(* IEC 61131-3 sources: daoli-st-library/DL_Motion (part 8) *)

(* ---- FB_DL_AxisOverspeedGuard.st ---- *)
(*
  FB_DL_AxisOverspeedGuard  —  轴超速守卫（速度窗 + 加速度窗双判据） / Axis overspeed guard with velocity and acceleration windows
  分类 Category : DL_Motion
  版本 Version  : 1.0.0
  来源 Source   : t2-4-s7motion — 运动守卫族零检索深化
  溯源 Origin   : clean-room 实现，未复制任何源码行
  功能 Function : 1) 速度判据：|fVelocity| > fVelMax 持续 tVelTo → 故障级 03AC 独立锁存；
                  2) 加速度判据：离散差分 fAccEst := |v - vPrev| / tSamp（采样周期单位
                  已在头注释声明 [mm/s 每秒]），fAccEst > fAccMax 持续 tAccTo →
                  故障级 03AD 独立锁存（R190 归因唯一：两成因各自独立码位与独立出口）；
                  3) 故障解除式全当拍量（R240 落地），逐 BOOL 标注见段 5；
                  4) 速度回窗置信息级 04AB，加速度回窗置 04AC，使能沿置 04AD。
  边界 Boundary : ① 组态闸：fVelMax <= 0、fAccMax <= 0、tSamp <= 0、两超时 <= 0 → 03AB 锁存；
                  ② 差分分母下限 1.0E-6 s 防除零（TIME_TO_LREAL 后钳位）；
                  ③ 速度窗下限语义：判据为绝对值上窗，无下窗（下限 0 显式化）；
                  ④ 无 GVL 依赖：纯引脚输入输出，无外部变量引用，无物理 IO 地址。
  依赖 Depends  : I_DL_MotionAxis（注入，不实例化）；Standard.library（TON / R_TRIG）
  码表 Error codes（Motion 段 0004，窗口 03AB~03AD / 04AB~04AD）:
    16#0004_03AB 故障级：组态非法（速度窗/加速度窗/采样周期/超时域非法），锁存至 bReset
    16#0004_03AC 故障级：超速锁存（速度窗判据），锁存至 bReset
    16#0004_03AD 故障级：加速度超窗锁存（加速度窗判据），锁存至 bReset
    16#0004_04AB 信息级：速度恢复正常沿（回速度窗内）
    16#0004_04AC 信息级：加速度恢复正常沿（回加速度窗内）
    16#0004_04AD 信息级：守卫使能沿（bEnable 上升沿）
  修订历史 Revision :
    2026-11-19  v1.0.0  R41 首版（批次 2 · 序号 5）
*)

FUNCTION_BLOCK FB_DL_AxisOverspeedGuard
VAR_INPUT
    fVelMax      : REAL := 1000.0;    // 速度窗上限绝对值 [mm/s]，域 > 0 / Velocity window upper bound
    fAccMax      : REAL := 5000.0;    // 加速度窗上限 [mm/s²]，域 > 0 / Acceleration window bound
    tSamp        : TIME := T#10MS;    // 差分采样周期 [ms]，域 > 0 / Differentiation sample period
    tVelTo       : TIME := T#100MS;   // 超速确认超时 [ms]，域 > 0 / Overspeed confirm timeout
    tAccTo       : TIME := T#100MS;   // 超加速度确认超时 [ms]，域 > 0 / Over-acceleration confirm timeout
    bEnable      : BOOL := FALSE;     // 守卫使能 [-] / Guard enable
    bReset       : BOOL := FALSE;     // 复位，上升沿清故障锁存 / Reset edge clears fault latch
END_VAR
VAR_IN_OUT
    iAxis        : I_DL_MotionAxis;   // 运动轴引用（注入，不实例化）/ Motion axis reference
END_VAR
VAR_OUTPUT
    fVelAct      : REAL;              // 速度出口镜像 [mm/s] / Velocity outlet mirror
    fAccEst      : REAL;              // 加速度离散估计 [mm/s²] / Discrete acceleration estimate
    bVelFault    : BOOL;              // 超速独立锁存出口 [-] / Overspeed latch outlet
    bAccFault    : BOOL;              // 超加速度独立锁存出口 [-] / Over-acceleration latch outlet
    bFault       : BOOL;              // 聚合故障标志 [-] / Aggregate fault flag
    bError       : BOOL;              // 故障级标志（与聚合锁存同源）/ Fault flag
    nErrId       : UDINT;             // 事件码，0 = 无事件 / Event code
END_VAR
VAR
    tonVelTo     : TON;               // 超速确认定时器，无条件周期刷新 / Overspeed confirm timer
    tonAccTo     : TON;               // 超加速度确认定时器，无条件周期刷新 / Over-acceleration confirm timer
    rtReset      : R_TRIG;            // 复位沿实例，无条件刷新 / Reset edge instance
    rtEn         : R_TRIG;            // 使能沿实例，无条件刷新 / Enable edge instance
    _fVel        : REAL;              // 速度当拍量 [mm/s] / Current-scan velocity
    _fVelPrev    : REAL;              // 上拍速度快照 [mm/s] / Previous-scan velocity snapshot
    _fSampSec    : REAL;              // 生效采样周期 [s] / Effective sample period in seconds
    _bVelLat     : BOOL;              // 超速锁存位（锁存量）/ Overspeed latch bit
    _bAccLat     : BOOL;              // 超加速度锁存位（锁存量）/ Over-acceleration latch bit
    _bCfgBad     : BOOL;              // 组态非法锁存位（锁存量）/ Config-fault latch bit
    _uFault      : UDINT;             // 故障码锁存（锁存量）/ Latched fault code
    _uInfo       : UDINT;             // 信息码，每拍重算 / Transient info code
    _bVelOkPrev  : BOOL;              // 上拍速度窗内镜像（恢复沿判据）/ Previous velocity-in-window mirror
    _bAccOkPrev  : BOOL;              // 上拍加速度窗内镜像（恢复沿判据）/ Previous acceleration-in-window mirror
END_VAR

(* —— 段 0：定时器与沿实例无条件周期刷新（禁置于 IF/CASE 内） —— *)
_fVel := iAxis.fVelocity;                              // 速度当拍量
_fSampSec := TIME_TO_LREAL(tSamp) * 1.0E-3;            // 采样周期换算秒 [s]
IF _fSampSec < 1.0E-6 THEN
    _fSampSec := 1.0E-6;            // 差分分母下限防除零（下限钳位）
END_IF
fAccEst := ABS(_fVel - _fVelPrev) / _fSampSec;         // 加速度离散估计（差分口径）
rtReset(CLK := bReset);                                // 复位沿（每拍必调）
rtEn(CLK := bEnable);                                  // 使能沿（每拍必调）
tonVelTo(IN := bEnable AND (ABS(_fVel) > fVelMax), PT := tVelTo);   // 超速确认（每拍必调）
tonAccTo(IN := bEnable AND (fAccEst > fAccMax), PT := tAccTo);      // 超加速度确认（每拍必调）

(* —— 段 1：单拍量预清零（锁存量 _uFault/_bVelLat/_bAccLat/_bCfgBad 不入清单，禁同拍抹除） —— *)
_uInfo := 16#0000_0000;             // 信息码每拍重算
nErrId := 16#0000_0000;             // 事件码缺省无事件

(* —— 段 2：复位沿 + 组态域闸（当拍量判据） —— *)
IF rtReset.Q THEN                   // rtReset.Q = 当拍量
    _bVelLat := FALSE;              // 清超速锁存位
    _bAccLat := FALSE;              // 清超加速度锁存位
    _bCfgBad := FALSE;              // 清组态锁存位
    _uFault := 16#0000_0000;        // 清故障锁存码
END_IF
IF (fVelMax <= 0.0) OR (fAccMax <= 0.0) OR (TIME_TO_DINT(tSamp) <= 0)
   OR (TIME_TO_DINT(tVelTo) <= 0) OR (TIME_TO_DINT(tAccTo) <= 0) THEN
    _uFault := 16#0004_03AB;        // 故障级：组态非法
    _bCfgBad := TRUE;
END_IF

(* —— 段 3：双判据独立锁存（R190：速度/加速度归因唯一，各走独立码位与出口） —— *)
IF (NOT _bCfgBad) AND tonVelTo.Q THEN
    _uFault := 16#0004_03AC;        // 故障级：超速锁存
    _bVelLat := TRUE;
END_IF
IF (NOT _bCfgBad) AND tonAccTo.Q THEN
    _uFault := 16#0004_03AD;        // 故障级：加速度超窗锁存
    _bAccLat := TRUE;
END_IF

(* —— 段 4：故障解除式（R240 落地，逐 BOOL 标注）：
     rtReset.Q = 当拍量；ABS(_fVel) <= fVelMax = 当拍量；fAccEst <= fAccMax = 当拍量。
     均不含锁存量（_bVelLat/_bAccLat），解除边真实可达。 —— *)
IF rtReset.Q AND (NOT _bCfgBad) AND (ABS(_fVel) <= fVelMax) AND (fAccEst <= fAccMax) THEN
    _bVelLat := FALSE;              // 清超速锁存位（锁存量，仅此当拍量解除沿可清）
    _bAccLat := FALSE;              // 清超加速度锁存位（锁存量，同上）
    _uFault := 16#0000_0000;        // 清故障锁存码（锁存量，同上唯一解除路径）
END_IF

(* —— 段 5：信息码派生（当拍量判据） —— *)
IF (NOT _bCfgBad) AND bEnable THEN
    IF (ABS(_fVel) <= fVelMax) AND (NOT _bVelOkPrev) THEN
        _uInfo := 16#0004_04AB;     // 信息级：速度恢复沿
    END_IF
    IF (fAccEst <= fAccMax) AND (NOT _bAccOkPrev) THEN
        _uInfo := 16#0004_04AC;     // 信息级：加速度恢复沿（覆盖速度恢复沿，后到优先）
    END_IF
END_IF
IF rtEn.Q THEN
    _uInfo := 16#0004_04AD;         // 信息级：使能沿（使能优先报告）
END_IF

(* —— 段 6：出口单点映射（名实同源；锁存码回放，禁同拍抹除） —— *)
fVelAct := _fVel;                   // 速度出口镜像
bVelFault := _bVelLat OR _bCfgBad;  // 超速独立出口（组态非法并入聚合安全侧）
bAccFault := _bAccLat OR _bCfgBad;  // 超加速度独立出口（同上）
bFault := _bVelLat OR _bAccLat OR _bCfgBad;     // 聚合故障
IF bFault THEN
    nErrId := _uFault;              // 故障锁存码回放
ELSE
    nErrId := _uInfo;               // 信息码
END_IF
bError := bFault;                   // 故障标志与聚合锁存同源
_bVelOkPrev := (ABS(_fVel) <= fVelMax);   // 速度恢复沿判据快照
_bAccOkPrev := (fAccEst <= fAccMax);      // 加速度恢复沿判据快照
_fVelPrev := _fVel;                 // 上拍速度快照（段末统一写）

END_FUNCTION_BLOCK

(* ---- FB_DL_AxisPowerOnSelfTest.st ---- *)
(*==============================================================================
 * 组件名称 (Component)  : FB_DL_AxisPowerOnSelfTest
 * 所属子库 (Sublibrary) : DL_Motion
 * 当前版本 (Version)    : 1.0.1
 * 兼容性   (Platform)   : CODESYS 3.5 / TwinCAT 3 / 汇川 InoProShop / Machine Expert
 *                         仅依赖 Standard.library（TON / R_TRIG），零厂商方言
 * 来源标签 (Source)     : t2-4-s7motion（上电自检序列语义，clean-room 编写）
 * 功能描述 (Function)   : 轴上电自检五步序检：驱动就绪 -> 编码器回读（位置有效性
 *                         + 速率合理性）-> 限位状态巡检（常开 / 常闭组态域闸）->
 *                         驱动故障字扫描 -> 结论锁存。任一步失败即中止并禁使能
 *                         放行：bTestOk 出口供 FB_DL_SingleAxis 使能链消费。
 * 家族纪律 (R31)        : 不自造轴状态枚举——本件只消费快照与反馈引脚
 *                         （bDriveReady / fEncPos / fEncRate / 限位位 / 故障字），
 *                         轴状态机归运动层接口 I_DL_MotionAxis，本件零轴状态定义。
 * 边界与语义披露 (Boundary disclosure) :
 *   1) 步序超时逐段 TON 断输入（R40 家族口径）：步切换拍计时器复位一次
 *      （IN 串「步激活 AND NOT 步更替」），各步共用同一 tStepTimeout。
 *   2) 结论锁存：bTestOk 只在结论相置位并保持；解除 = 复位沿 AND 驱动就绪在位
 *      （终审两式：解除式可达，验收向量「复位沿 + 驱动就绪 -> 可重测」）。
 *   3) 限位组态域闸：nLimitMode 仅 0（常开）/ 1（常闭）合法，其余组态级故障；
 *      常闭口径下反馈 TRUE = 未压（健康），常开口径下反馈 TRUE = 被压。
 *   4) 上电即被压的限位按自检失败处置（轴未能验证自由行程，放行风险不可接受）。
 *   5) 编码器回读判据：位置 / 速率非有限（自反 + 差自减双判）或 |速率| 超
 *      fRateMax 均判步 2 失败（验收向量：回读 NaN -> 步 2 中止 bTestOk FALSE 置码）。
 *   6) 通用组态（速率上限 / 步超时）非法独立码位，与限位组态成因互异（R190）。
 * 故障码表 (Error codes) :
 *   16#0004_0363 [故障级] 步序超时（当前步 tStepTimeout 未达成）
 *                 反证：超时中止与「判据失败中止」eFault 输出组合相同，成因必须码位互异。
 *   16#0004_0364 [故障级] 编码器回读非法（位置 / 速率非有限或速率超合理域）
 *                 反证：步 2 中止与其它步中止输出组合相似，码位是唯一成因出口。
 *   16#0004_0365 [故障级] 限位组态模式非法（nLimitMode 非 0 / 1）
 *                 反证：限位步失败与编码器步失败输出组合相似，码位互异（R190）。
 *   16#0004_0366 [故障级] 上电限位被压（按生效接线口径判），自由行程未验证
 *                 反证：与组态非法同相中止但成因互异，码位独立。
 *   16#0004_0367 [故障级] 驱动故障字非零
 *                 反证：驱动故障字中止与编码器 / 限位 / 超时中止输出组合相似，成因互异码位独立。
 *   16#0004_0368 [故障级] 通用组态非法（速率上限 / 步超时域），拒绝启动
 *                 反证：拒绝启动与「未按触发」输出组合相同，码位唯一可见。
 * 码位总账 (Code ledger) : 16#0004_0363 / 0364 / 0365 / 0366 / 0367 / 0368 用
 * 依赖     (Depends)    : 无 DL_ 内部依赖；Standard.library: TON / R_TRIG
 * 红线自检 (Redline)    : R1 ✓ 零全局变量与 VAR_EXTERNAL ｜ R2 ✓ 零 %I/%Q 物理地址
 *                         R3 ✓ 纯 IEC 61131-3 ｜ R4 ✓ 非有限双判 / 域闸全枚举 / 码位 R45 配对
 *                         R5 ✓ 全变量中英双语同行注释 ｜ R6 ✓ 七态 ENUM + CASE + ELSE 兜底
 *                         R7 ✓ 三沿一计时主体最前部无条件刷新
 * 修订历史 (Revision)   :
 *   2026-11-22  v1.0.0  首版入库（R68 构建轮 · 批 3 · 目标 16）
 *   2026-11-22  v1.0.1  终审就地修①：组态锁存解除路径可达化（原 bCfgLatch 全文件零清零 -> 自检永久不可重测）
 *============================================================================*)

(*-----------------------------------------------------------------------------
 * 枚举: E_DL_SelfTestStep（归属 DL_Motion，与 FB_DL_AxisPowerOnSelfTest 同文件）
 * 说明: 本枚举是「自检步序」不是「轴状态」——轴状态归运动层接口（R31 家族纪律）。
 *----------------------------------------------------------------------------*)
TYPE E_DL_SelfTestStep :
(
    eIdle        := 0,    // 待触发：结论保持 / Idle, conclusion held
    eStDrive     := 10,   // 步 1：驱动就绪确认 / Step 1, drive ready
    eStEncoder   := 20,   // 步 2：编码器回读校验 / Step 2, encoder readback
    eStLimits    := 30,   // 步 3：限位状态巡检 / Step 3, limit switch patrol
    eStDriveWord := 40,   // 步 4：驱动故障字扫描 / Step 4, drive fault word scan
    eStConclude  := 50,   // 步 5：结论锁存 / Step 5, conclusion latch
    eFault       := 99    // 自检失败锁存：禁使能放行 / Self-test failed, enable release denied
);
END_TYPE

(*==============================================================================
 * 功能块: FB_DL_AxisPowerOnSelfTest
 * 调用约定: 每个扫描周期无条件调用一次；快照引脚须每拍刷新注入。
 *============================================================================*)
FUNCTION_BLOCK FB_DL_AxisPowerOnSelfTest
VAR_INPUT
    bTestTrig    : BOOL;                  // 自检触发（上升沿受理）/ Self-test trigger, rising edge
    bDriveReady  : BOOL;                  // 驱动就绪快照 / Drive ready snapshot
    fEncPos      : LREAL;                 // 编码器位置回读 [mm] / Encoder position readback [mm]
    fEncRate     : LREAL;                 // 编码器速率回读 [mm/s] / Encoder rate readback [mm per s]
    fRateMax     : LREAL := 100.0;        // 速率合理上限 [mm/s] / Plausible rate ceiling [mm per s]
    bLimitPosFb  : BOOL;                  // 正限位状态反馈（原始，TRUE = 电气有效）/ Positive limit feedback, raw
    bLimitNegFb  : BOOL;                  // 负限位状态反馈（原始）/ Negative limit feedback, raw
    nLimitMode   : INT   := 0;            // 限位接线模式：0 = 常开，1 = 常闭 / Wiring mode, 0 NO 1 NC
    uDriveFaultWord : WORD;               // 驱动故障字 / Drive fault word
    tStepTimeout : TIME  := T#2S;         // 单步超时 [s] / Step timeout [s]
    bEnable      : BOOL  := TRUE;         // 使能 / Enable
    bReset       : BOOL;                  // 上升沿：清结论与故障锁存（须驱动就绪在位）/ Rising edge: clear, drive ready required
END_VAR
VAR_OUTPUT
    bTestOk    : BOOL;                   // 自检结论：TRUE = 通过（锁存至复位 / 新测）/ Test passed, latched
    bTestDone  : BOOL;                   // 结论已出（通过或失败）/ Conclusion available
    bError     : BOOL;                   // 故障标志（自检失败 / 组态锁存归并）/ Fault flag merged
    uErrorId   : UDINT;                  // 故障码，0 = 无故障 / Error code, 0 = none
    eState     : E_DL_SelfTestStep;      // 当前步序（供 HMI 诊断）/ Current step for HMI diagnosis
END_VAR
VAR
    fbTrigTrig  : R_TRIG;                // 触发沿检测实例 / Trigger edge detector
    fbTrigReset : R_TRIG;                // 复位沿检测实例 / Reset edge detector
    tonStep     : TON;                   // 单步超时计时实例 / Step timeout timer
    eStateInt   : E_DL_SelfTestStep;     // 主状态机内部当前态 / Internal state machine state
    eStepPrev   : E_DL_SelfTestStep;     // 上拍步序快照（步更替判据）/ Previous step snapshot
    bStepActive : BOOL;                  // 当前步处于计时激活域 / Current step in the timed set
    bStepNew    : BOOL;                  // 本拍发生步更替（计时复位点）/ Step changed this scan
    bLimPosTrip : BOOL;                  // 按接线口径判的正限位被压 / Positive limit tripped per wiring
    bLimNegTrip : BOOL;                  // 负限位被压 / Negative limit tripped
    bEncBad     : BOOL;                  // 编码器回读非法 / Encoder readback illegal
    bCfgBad     : BOOL;                  // 本拍通用组态非法 / General config illegal
    bCfgLatch   : BOOL;                  // 通用组态锁存 / General config latch
    bModeBad    : BOOL;                  // 限位接线模式非法 / Wiring mode illegal
    bPassedInt  : BOOL;                  // 通过结论锁存内部副本 / Internal passed latch
    bDoneInt    : BOOL;                  // 结论已出锁存内部副本 / Internal done latch
    bErrorInt   : BOOL;                  // 本拍故障置位累加（出口归并）/ Fault set accumulator
    bFirstScan  : BOOL := TRUE;          // 上电首扫标志 / First-scan flag
END_VAR
VAR CONSTANT
    DL_ST_FIN_LIM   : LREAL := 1.0E30;   // LREAL 有限幅值判界 / LREAL finiteness bound
    DL_ST_MODE_NO   : INT   := 0;        // 常开接线模式号 / Normally-open mode id
    DL_ST_MODE_NC   : INT   := 1;        // 常闭接线模式号 / Normally-closed mode id
END_VAR

(*------------------------------------------------------------------------------
 * 段 1｜无条件刷新区（红线 R7）：二沿一计时主体最前部
 *      Unconditional refresh: two edges and one timer at the very top
 *      步更替拍计时复位一次（IN 串「步激活 AND NOT 步更替」，逐段断输入 R40）
 *-----------------------------------------------------------------------------*)
fbTrigTrig(CLK := bTestTrig);
fbTrigReset(CLK := bReset);

bStepNew := (eStateInt <> eStepPrev);

bStepActive := (eStateInt = E_DL_SelfTestStep.eStDrive)
               OR (eStateInt = E_DL_SelfTestStep.eStEncoder)
               OR (eStateInt = E_DL_SelfTestStep.eStLimits)
               OR (eStateInt = E_DL_SelfTestStep.eStDriveWord);

tonStep(IN := bStepActive AND (NOT bStepNew), PT := tStepTimeout);

(*------------------------------------------------------------------------------
 * 段 2｜上电首扫：结论与状态落安全侧（未测 = 不放行）
 *      First-scan init: conclusion to the safe side, untested means no release
 *-----------------------------------------------------------------------------*)
IF bFirstScan THEN
    eStateInt  := E_DL_SelfTestStep.eIdle;
    eStepPrev  := eStateInt;
    bPassedInt := FALSE;
    bDoneInt   := FALSE;
    bFirstScan := FALSE;
END_IF

(*------------------------------------------------------------------------------
 * 段 3｜每拍预清（FB32-1）：单拍标志，禁入锁存 / 快照
 *      Per-scan preset: single-scan flags only
 *-----------------------------------------------------------------------------*)
bErrorInt := FALSE;

(*------------------------------------------------------------------------------
 * 段 4｜组态域闸（R151 全枚举）：通用组态 + 限位接线模式（独立成因独立码 R190）
 *      Config gates: general config plus the wiring mode, distinct codes
 *      解除路径（R152 自证）：复位沿 AND 驱动就绪 AND 组态改对
 *-----------------------------------------------------------------------------*)
bCfgBad := (fRateMax <= 0.0) OR (fRateMax <> fRateMax) OR (tStepTimeout <= T#0S);
bModeBad := (nLimitMode <> DL_ST_MODE_NO) AND (nLimitMode <> DL_ST_MODE_NC);

IF bCfgBad THEN
    bCfgLatch := TRUE;
    uErrorId  := 16#0004_0368;    // 故障级：通用组态非法 / Fault: general config illegal
    bErrorInt := TRUE;
END_IF

(* 终审就地修 v1.0.1（R68）：解除路径（R152 自证可达）——复位沿 AND 组态非法条件
 * 全部消失即清锁存。原实现把锁存清零只写在 eFault 相分支，而组态闸置锁存后
 * 并不迁相至 eFault（只回 eIdle / 驻留），eFault 相不可达 -> 锁存永不可解，
 * 组件保护/监视功能一次性永久失效直至 PLC 重启（终审两式①）。
 * Clear path made provably reachable: reset edge with the illegal config gone. *)
IF fbTrigReset.Q AND (NOT bCfgBad) THEN
    bCfgLatch := FALSE;           // 锁存解除 / Latch cleared
    uErrorId  := 16#0000_0000;    // 码位随解除归零 / Code cleared with the latch
END_IF

(*------------------------------------------------------------------------------
 * 段 5｜限位接线口径换算（步 3 判据核）：常闭反馈 TRUE = 健康，常开反馈 TRUE = 被压
 *      Limit wiring translation: NC TRUE = healthy, NO TRUE = tripped
 *-----------------------------------------------------------------------------*)
IF nLimitMode = DL_ST_MODE_NC THEN
    bLimPosTrip := NOT bLimitPosFb;      // 常闭：未反馈即被压 / NC: no feedback means tripped
    bLimNegTrip := NOT bLimitNegFb;
ELSE
    bLimPosTrip := bLimitPosFb;          // 常开：有反馈即被压 / NO: feedback means tripped
    bLimNegTrip := bLimitNegFb;
END_IF

(*------------------------------------------------------------------------------
 * 段 6｜主状态机（红线 R6）：ENUM + CASE + ELSE 兜底
 *      Main state machine with the mandatory ELSE fallback
 *-----------------------------------------------------------------------------*)
CASE eStateInt OF

    E_DL_SelfTestStep.eIdle:
        IF bCfgLatch OR (NOT bEnable) THEN
            (* 组态 / 失能驻留：结论保持不放行 / Dwell, conclusion held, no release *)
        ELSIF fbTrigTrig.Q AND bModeBad THEN
            (* 触发但接线组态非法：拒绝启动并落组态码（不允许带病起测） *)
            (* Trigger with illegal wiring: refused with the mode code *)
            uErrorId  := 16#0004_0365;
            bErrorInt := TRUE;
        ELSIF fbTrigTrig.Q THEN
            bPassedInt := FALSE;     // 新测清旧结论 / New test clears the old verdict
            bDoneInt   := FALSE;
            eStateInt  := E_DL_SelfTestStep.eStDrive;
        END_IF

    E_DL_SelfTestStep.eStDrive:
        IF tonStep.Q THEN
            eStateInt := E_DL_SelfTestStep.eFault;   // 步 1 超时 / Step 1 timeout
            uErrorId  := 16#0004_0363;
            bErrorInt := TRUE;
        ELSIF bDriveReady THEN
            eStateInt := E_DL_SelfTestStep.eStEncoder;   // 就绪进步 2 / Ready, to step 2
        END_IF

    E_DL_SelfTestStep.eStEncoder:
        bEncBad := (fEncPos <> fEncPos)
                   OR ((fEncPos - fEncPos) <> (fEncPos - fEncPos))
                   OR (ABS(fEncPos) >= DL_ST_FIN_LIM)
                   OR (fEncRate <> fEncRate)
                   OR ((fEncRate - fEncRate) <> (fEncRate - fEncRate))
                   OR (ABS(fEncRate) >= DL_ST_FIN_LIM)
                   OR (ABS(fEncRate) > fRateMax);
        IF tonStep.Q THEN
            eStateInt := E_DL_SelfTestStep.eFault;
            uErrorId  := 16#0004_0363;
            bErrorInt := TRUE;
        ELSIF bEncBad THEN
            eStateInt := E_DL_SelfTestStep.eFault;   // 步 2 中止（验收向量：NaN 回读）/ Step 2 abort
            uErrorId  := 16#0004_0364;
            bErrorInt := TRUE;
        ELSE
            eStateInt := E_DL_SelfTestStep.eStLimits;    // 回读合法进步 3 / Valid, to step 3
        END_IF

    E_DL_SelfTestStep.eStLimits:
        IF tonStep.Q THEN
            eStateInt := E_DL_SelfTestStep.eFault;
            uErrorId  := 16#0004_0363;
            bErrorInt := TRUE;
        ELSIF bModeBad THEN
            eStateInt := E_DL_SelfTestStep.eFault;   // 接线组态非法 / Wiring mode illegal
            uErrorId  := 16#0004_0365;
            bErrorInt := TRUE;
        ELSIF bLimPosTrip OR bLimNegTrip THEN
            eStateInt := E_DL_SelfTestStep.eFault;   // 上电限位被压 / Limit tripped at power-on
            uErrorId  := 16#0004_0366;
            bErrorInt := TRUE;
        ELSE
            eStateInt := E_DL_SelfTestStep.eStDriveWord; // 限位健康进步 4 / Healthy, to step 4
        END_IF

    E_DL_SelfTestStep.eStDriveWord:
        IF tonStep.Q THEN
            eStateInt := E_DL_SelfTestStep.eFault;
            uErrorId  := 16#0004_0363;
            bErrorInt := TRUE;
        ELSIF uDriveFaultWord <> 16#0000 THEN
            eStateInt := E_DL_SelfTestStep.eFault;   // 驱动故障字非零 / Fault word nonzero
            uErrorId  := 16#0004_0367;
            bErrorInt := TRUE;
        ELSE
            eStateInt := E_DL_SelfTestStep.eStConclude;  // 故障字干净进步 5 / Clean, to step 5
        END_IF

    E_DL_SelfTestStep.eStConclude:
        bPassedInt := TRUE;          // 五步全过：通过结论锁存 / All steps pass: latch the verdict
        bDoneInt   := TRUE;
        eStateInt  := E_DL_SelfTestStep.eIdle;

    E_DL_SelfTestStep.eFault:
        bDoneInt := TRUE;            // 失败结论已出 / Failure verdict available
        (* 解除路径（R152 自证可达）：复位沿 AND 驱动就绪在位 AND 组态改对（可重测） *)
        IF fbTrigReset.Q AND bDriveReady AND (NOT bCfgBad) AND (NOT bModeBad) THEN
            uErrorId  := 16#0000_0000;
            eStateInt := E_DL_SelfTestStep.eIdle;
        END_IF

    ELSE
        (* 非法状态拦截：迁兜底态（复用组态段码位） *)
        eStateInt := E_DL_SelfTestStep.eFault;
        uErrorId  := 16#0004_0368;
        bErrorInt := TRUE;

END_CASE;

(*------------------------------------------------------------------------------
 * 段 7｜步序快照（主体末行，R45 累计定时器留上拍快照口径的同族纪律）
 *      Step snapshot at the body tail
 *-----------------------------------------------------------------------------*)
eStepPrev := eStateInt;

(*------------------------------------------------------------------------------
 * 段 8｜输出单一出口（范式 P-05）：结论只由锁存派生
 *      Single output exit: the verdict derives from the latch only
 *      测试未通过时 bTestOk 恒 FALSE（无恒假锁存——结论只写 TRUE 一次）
 *-----------------------------------------------------------------------------*)
bTestOk   := bPassedInt;
bTestDone := bDoneInt;
bError    := bErrorInt OR (eStateInt = E_DL_SelfTestStep.eFault);
eState    := eStateInt;
END_FUNCTION_BLOCK

(* ---- FB_DL_AxisProbeMeasCycle.st ---- *)
(*
  ==================================================================
  组件名 Component  : FB_DL_AxisProbeMeasCycle
  分类   Category   : DL_Motion
  复杂度 Complexity  : cx5
  版本   Version    : 1.0.0
  功能   Purpose    : 探针测量循环。相位机 eIdle → eFastApproach → eProbeLatch →
                      eRetract → eSettle → eRecord → eDone / eFault；快进 - 慢探
                      两段速度；探针触发用 R_TRIG 边沿锁存（锁存值用于记录，
                      禁与实时镜像混用）；超行程保护；nRepeat 次重复测量后做
                      离散度判据（max - min 对容差），超差判 eScatterHigh。
  来源   Source     : t2-2-lbp（与 FB_DL_MarkPositionLatch 分工：锁存原子 vs 完整测量循环）
  溯源   Origin     : IEC 61131-3 标准语义的道莅防御性实现；趋近 - 触发锁存 - 回退 -
                      评价测量循环为通用测量语义，clean-room 自研实现，未复制任何
                      闭源代码行。
  平台   Platform   : 纯 IEC 61131-3（TON / R_TRIG / ARRAY / LREAL，无私有库）
  作者   Author     : 道莅代码库 · PLC 编程专家（R56）
  ------------------------------------------------------------------
  同拍多窗说明（R100）：四个窗互斥 —— 每窗 IN 串「本相」闸，任一时刻只有一个窗
                      在计时，无同拍双窗配比约束。
  边界 Boundary     :
                      一 本件只出速度命令与测量结论，不驱动轴本体、不解算几何尺寸
                         （属主边界）；
                      二 锁存纪律：_fMeasPos 只在触发沿那一拍由 fPosAct 写入一次，
                         其后评价一律用锁存值（R33 锁存副本与实时镜像不混用）；
                      三 相级看门狗使能只用相驻留本身（R145）；
                      四 故障锁存解除路径 = bReset 上升沿（唯一路径，R188）；
                      五 无全局变量、无外部变量声明、无物理地址寻址。
  输出契约 Output contract:
                      fVelCmd 为速度命令（快进 / 慢探 / 回退三档）；fMeasPos 为
                      nRepeat 次均值；bMeasValid 为单拍脉冲（R187 两段式）；
                      eFault 为锁存回放；ePhaseBad 为非法相位兜底专用成员（R128）。
  修订记录 Revision  :
    2026-11-20  v1.0.0  R56 首版（批 4 · 序号 19）
  ==================================================================
*)

TYPE E_DL_ApcPhase :
(
    eIdle         := 0,  // 空闲：等启动沿 / idle, waiting for the start edge
    eFastApproach := 10, // 快进：高速趋近到慢探起点 / fast approach, high speed to the slow start
    eProbeLatch   := 20, // 慢探：低速探触发并锁存 / probe latch, low speed to the trigger with a latch
    eRetract      := 30, // 回退：退回安全距 / retract, back to the safe distance
    eSettle       := 40, // 稳定：驻留稳定窗 / settle, the dwell window
    eRecord       := 50, // 记录：样本入环并评价 / record, the sample enters the ring and the verdict runs
    eDone         := 60, // 完成：结论驻留 / done, the verdict holds
    eFault        := 90  // 故障：成因锁存 / fault, the cause is latched
);
END_TYPE

TYPE E_DL_ApcFault :
(
    eNone       := 0, // 无成因 / no cause
    eNoTrigger  := 1, // 越程内未触发（故障级，与 bError 配对）/ no trigger inside the travel limit, fault grade paired with bError
    eOverTravel := 2, // 超行程保护（故障级，与 bError 配对）/ the overtravel protection, fault grade paired with bError
    eScatterHigh:= 3, // 重复测量离散度超差（故障级，与 bError 配对）/ the scatter of the repeats is over the tolerance, fault grade paired with bError
    eSensorBad  := 4, // 位置非有限或组态非法（故障级，与 bError 配对）/ the position is non finite or the config illegal, fault grade paired with bError
    ePhaseBad   := 5  // 非法相位兜底（故障级，与 bError 配对）/ illegal phase fallback, fault grade paired with bError
);
END_TYPE

FUNCTION_BLOCK FB_DL_AxisProbeMeasCycle
VAR_INPUT
    bEnable     : BOOL := TRUE;    // 使能，失能时停循环回空闲 [-] / enable, the cycle stops when disabled
    bReset      : BOOL := FALSE;   // 复位上升沿清故障锁存与样本环 [-] / reset rising edge clears the latch and the sample ring
    bStart      : BOOL := FALSE;   // 测量启动脉冲，上升沿受理 [-] / the measurement start pulse, accepted on the rising edge
    bAbort      : BOOL := FALSE;   // 中止（电平），任何中间态回空闲 [-] / the abort level, any middle phase returns to idle
    fPosAct     : LREAL := 0.0;    // 轴实际位置 [位置单位] / the actual axis position [position unit]
    bProbeTrig  : BOOL := FALSE;   // 探针触发信号 [-] / the probe trigger signal
    fTargetPos  : LREAL := 100.0;  // 目标标称位置 [位置单位] / the nominal target position [position unit]
    fSlowStart  : LREAL := 90.0;   // 慢探起点（快进切换位）[位置单位] / the slow probe start [position unit]
    fBackDist   : LREAL := 5.0;    // 回退安全距 [位置单位]，域 大于零 / the retract safe distance [position unit], domain above zero
    fOverTravel : LREAL := 2.0;    // 超行程容限（越程即故障 / 未触发判据）[位置单位]，域 大于零 / the overtravel tolerance [position unit], domain above zero
    fScatterTol : LREAL := 0.01;   // 离散度容差 [位置单位]，域 大于零 / the scatter tolerance [position unit], domain above zero
    nRepeat     : INT := 3;        // 重复测量次数 [次]，域 1..20 / the repeat count [count], domain one to twenty
    fVelFast    : LREAL := 500.0;  // 快进速度 [位置单位每秒] / the fast approach velocity [position unit per second]
    fVelSlow    : LREAL := 20.0;   // 慢探速度 [位置单位每秒]，域 小于快进 / the slow probe velocity, below the fast one
    tFastTo     : TIME := T#10S;   // 快进超时窗 [毫秒] / the fast approach timeout [millisecond]
    tProbeTo    : TIME := T#10S;   // 慢探超时窗 [毫秒] / the probe timeout [millisecond]
    tRetractTo  : TIME := T#5S;    // 回退超时窗 [毫秒] / the retract timeout [millisecond]
    tSettle     : TIME := T#200MS; // 稳定驻留窗 [毫秒] / the settle dwell window [millisecond]
END_VAR
VAR_OUTPUT
    fVelCmd   : LREAL := 0.0;   // 速度命令（快进 / 慢探 / 回退三档）[位置单位每秒] / the velocity command, three gears [position unit per second]
    fMeasPos  : LREAL := 0.0;   // 测量结论（nRepeat 次均值）[位置单位] / the measurement verdict, the mean of the repeats [position unit]
    bMeasValid: BOOL := FALSE;  // 测量有效单拍脉冲 [-] / the measurement valid single shot pulse
    nMeasCnt  : INT := 0;       // 已完成测量次数 [次] / the completed measurement count [count]
    ePhase    : E_DL_ApcPhase := E_DL_ApcPhase.eIdle; // 相位出口 [枚举] / phase outlet [enum]
    eFault    : E_DL_ApcFault := E_DL_ApcFault.eNone; // 成因出口，锁存回放 [枚举] / cause outlet replayed from the latch [enum]
    bError    : BOOL := FALSE;  // 故障锁存标志 [-] / fault latch flag
END_VAR
VAR
    rtStart  : R_TRIG; // 启动沿检测，段 0 无条件刷新 / start edge, refreshed unconditionally in segment zero
    rtProbe  : R_TRIG; // 探针触发沿检测，段 0 无条件刷新 / the probe trigger edge, refreshed unconditionally in segment zero
    rtReset  : R_TRIG; // 复位沿检测，段 0 无条件刷新 / reset edge, refreshed unconditionally in segment zero
    tonFast  : TON;    // 快进超时窗，段 0 无条件刷新 / the fast timeout window, refreshed unconditionally
    tonProbe : TON;    // 慢探超时窗，段 0 无条件刷新 / the probe timeout window, refreshed unconditionally
    tonRetr  : TON;    // 回退超时窗，段 0 无条件刷新 / the retract timeout window, refreshed unconditionally
    tonSettle: TON;    // 稳定驻留窗，段 0 无条件刷新 / the settle dwell window, refreshed unconditionally
    _ePhase  : E_DL_ApcPhase := E_DL_ApcPhase.eIdle; // 内部相位，CASE 唯一写入目标 / internal phase, the only CASE write target
    _eFaulC  : E_DL_ApcFault := E_DL_ApcFault.eNone; // 故障级成因，锁存至复位沿 / fault cause, latched until the reset edge
    _bFault  : BOOL := FALSE; // 故障锁存位 [-] / fault latch bit
    _bInit   : BOOL := FALSE; // 首扫初始化完成标志（R310）/ first scan initialisation flag
    _bDoneInt: BOOL := FALSE; // 有效脉冲内部位，统一出口映射 / internal valid bit, mapped at the unified outlet
    _bInOk   : BOOL := FALSE; // 位置有限 [-] / the position is finite
    _bCfgOk  : BOOL := FALSE; // 组态参数域内 [-] / the configuration is inside the domain
    _fLatch  : LREAL := 0.0;  // 触发沿锁存位置（评价唯一来源）[位置单位] / the latched position at the trigger edge, the only evaluation source
    _fMax    : LREAL := 0.0;  // 样本最大值 [位置单位] / the sample maximum [position unit]
    _fMin    : LREAL := 0.0;  // 样本最小值 [位置单位] / the sample minimum [position unit]
    _fSum    : LREAL := 0.0;  // 样本和 [位置单位] / the sample sum [position unit]
    _nRepeat : INT := 3;      // 钳定后的重复次数 [次] / the clamped repeat count [count]
    _nCnt    : INT := 0;      // 已收样本数 [个] / the collected sample count [count]
    _nI      : INT := 1;      // 环窗遍历游标 [槽号] / the ring traversal cursor
    _nGuard  : INT := 0;      // 遍历守护计数 [次] / the traversal guard [count]
    _anMeas  : ARRAY[1..20] OF LREAL := [20(0.0)]; // 样本环（时间序追加，无回绕需求）[位置单位] / the sample ring appended in time order [position unit]
END_VAR

// 段 0｜定时器与沿检测无条件周期刷新（禁入分支），IN 只串相位闸与故障闸（FB50-1）/ segment 0, unconditional refresh, no instance call inside a branch
rtStart(CLK := bStart); // 启动沿 / the start edge
rtProbe(CLK := bProbeTrig); // 探针触发沿 / the probe trigger edge
rtReset(CLK := bReset); // 复位沿 / the reset edge
tonFast(IN := (_ePhase = E_DL_ApcPhase.eFastApproach) AND (NOT _bFault), PT := tFastTo); // 快进超时窗 / the fast timeout window
tonProbe(IN := (_ePhase = E_DL_ApcPhase.eProbeLatch) AND (NOT _bFault), PT := tProbeTo); // 慢探超时窗 / the probe timeout window
tonRetr(IN := (_ePhase = E_DL_ApcPhase.eRetract) AND (NOT _bFault), PT := tRetractTo); // 回退超时窗 / the retract timeout window
tonSettle(IN := (_ePhase = E_DL_ApcPhase.eSettle) AND (NOT _bFault), PT := tSettle); // 稳定驻留窗 / the settle dwell window

// 段 1｜首扫初始化（R310）/ segment 1, first scan initialisation
IF NOT _bInit THEN // 首扫一拍 / the very first scan
    _bInit := TRUE; // 置首扫完成标志 / raise the first scan flag
    _ePhase := E_DL_ApcPhase.eIdle; // 相位从空闲起步 / the phase starts from idle
    _eFaulC := E_DL_ApcFault.eNone; // 故障级成因清零 / clear the fault cause
    _bFault := FALSE; // 故障锁存清零 / clear the fault latch
    _nCnt := 0; // 样本数清零 / clear the sample count
END_IF

// 段 2｜复位沿作用域：清锁存 / 迁相位 / 清样本环与计数（三项逐项声明）/ segment 2, reset edge scope declared item by item
IF rtReset.Q THEN // 复位沿 / the reset edge
    _bFault := FALSE; // 作用域一：清故障锁存 / scope one, clear the fault latch
    _eFaulC := E_DL_ApcFault.eNone; // 作用域一：清故障级成因 / scope one, clear the fault cause
    _ePhase := E_DL_ApcPhase.eIdle; // 作用域二：迁回空闲相 / scope two, migrate back to idle
    _nCnt := 0; // 作用域三：清样本计数 / scope three, clear the sample count
    fVelCmd := 0.0; // 作用域三：速度命令归零 / scope three, the velocity command zeroes
END_IF

// 段 3｜组态与输入域闸（R151 全覆盖）/ segment 3, the configuration and input domain gates
_bInOk := (fPosAct = fPosAct) AND ((fPosAct - fPosAct) = (fPosAct - fPosAct)); // 位置有限性 / the position finiteness
_bCfgOk := (fBackDist > 0.0) AND (fBackDist = fBackDist) AND (fOverTravel > 0.0) AND (fOverTravel = fOverTravel) AND (fScatterTol > 0.0) AND (fScatterTol = fScatterTol) AND (fVelFast > 0.0) AND (fVelFast = fVelFast) AND (fVelSlow > 0.0) AND (fVelSlow < fVelFast) AND (fVelSlow = fVelSlow) AND (tFastTo > T#0S) AND (tProbeTo > T#0S) AND (tRetractTo > T#0S) AND (tSettle > T#0S); // 组态参数域判定 / the configuration domain verdict
_nRepeat := nRepeat; // 重复次数直通 / the repeat count passes through
IF _nRepeat < 1 THEN // 下越域 / below the floor
    _nRepeat := 1; // 回钳到一 / clamp to one
ELSIF _nRepeat > 20 THEN // 上越域 / above the ceiling
    _nRepeat := 20; // 回钳到二十 / clamp to twenty
END_IF
IF (NOT _bInOk) OR (NOT _bCfgOk) THEN // 位置非有限或组态非法 / a void position or an illegal configuration
    IF NOT _bFault THEN // 未锁存才迁移（防同拍抹除）/ migrate only while unlatched
        _bFault := TRUE; // 置故障锁存 / raise the fault latch
        _eFaulC := E_DL_ApcFault.eSensorBad; // 故障级成因（R45 配对 bError）/ the fault cause paired with bError
        _ePhase := E_DL_ApcPhase.eFault; // 迁故障相 / migrate to the fault phase
    END_IF
END_IF

// 段 4｜相位机：ENUM + CASE，含 ELSE 非法相位兜底（R128）/ segment 4, the phase machine with an ELSE fallback
CASE _ePhase OF
E_DL_ApcPhase.eIdle: // 空闲相：等启动沿 / the idle phase, waiting for the start edge
    fVelCmd := 0.0; // 速度命令归零 / the velocity command zeroes
    IF bEnable AND (NOT _bFault) AND (NOT bAbort) AND rtStart.Q THEN // 启动沿受理 / the start edge is accepted
        _nCnt := 0; // 样本数清零（新测量批次）/ clear the sample count for a fresh batch
        _ePhase := E_DL_ApcPhase.eFastApproach; // 迁快进相 / migrate to the fast approach phase
    END_IF

E_DL_ApcPhase.eFastApproach: // 快进相：高速趋近（退出条件 ≥2：到慢探起点 / 超时 / 越程 / 中止 / 失能，R98）/ the fast approach phase with at least two exit conditions
    fVelCmd := fVelFast; // 快进速度命令 / the fast velocity command
    IF (NOT bEnable) OR bAbort THEN // 失能或中止 / disabled or aborting
        _ePhase := E_DL_ApcPhase.eIdle; // 回空闲相 / back to idle
    ELSIF NOT _bInOk THEN // 位置非有限 / the position went void
        _bFault := TRUE; // 置故障锁存 / raise the fault latch
        _eFaulC := E_DL_ApcFault.eSensorBad; // 故障级成因（R45 配对 bError）/ the fault cause paired with bError
        _ePhase := E_DL_ApcPhase.eFault; // 迁故障相 / migrate to the fault phase
    ELSIF fPosAct > fTargetPos + fOverTravel THEN // 超行程保护（R146 安全侧立即终止）/ the overtravel protection, an immediate safe side stop
        _bFault := TRUE; // 置故障锁存 / raise the fault latch
        _eFaulC := E_DL_ApcFault.eOverTravel; // 故障级成因（R45 配对 bError）/ the fault cause paired with bError
        _ePhase := E_DL_ApcPhase.eFault; // 迁故障相 / migrate to the fault phase
    ELSIF fPosAct >= fSlowStart THEN // 到慢探起点 / the slow start is reached
        _ePhase := E_DL_ApcPhase.eProbeLatch; // 迁慢探相 / migrate to the probe latch phase
    ELSIF tonFast.Q THEN // 快进超时 / the fast approach timed out
        _bFault := TRUE; // 置故障锁存 / raise the fault latch
        _eFaulC := E_DL_ApcFault.eNoTrigger; // 故障级成因（R45 配对 bError，快进未达判慢探必不触发）/ the fault cause paired with bError
        _ePhase := E_DL_ApcPhase.eFault; // 迁故障相 / migrate to the fault phase
    END_IF

E_DL_ApcPhase.eProbeLatch: // 慢探相：低速探触发并锁存 / the probe latch phase, the low speed trigger with the latch
    fVelCmd := fVelSlow; // 慢探速度命令 / the slow velocity command
    IF (NOT bEnable) OR bAbort THEN // 失能或中止 / disabled or aborting
        _ePhase := E_DL_ApcPhase.eIdle; // 回空闲相 / back to idle
    ELSIF NOT _bInOk THEN // 位置非有限 / the position went void
        _bFault := TRUE; // 置故障锁存 / raise the fault latch
        _eFaulC := E_DL_ApcFault.eSensorBad; // 故障级成因（R45 配对 bError）/ the fault cause paired with bError
        _ePhase := E_DL_ApcPhase.eFault; // 迁故障相 / migrate to the fault phase
    ELSIF fPosAct > fTargetPos + fOverTravel THEN // 越程未触发（超行程判据复用，R146 方向一致）/ past the limit without a trigger
        _bFault := TRUE; // 置故障锁存 / raise the fault latch
        _eFaulC := E_DL_ApcFault.eNoTrigger; // 故障级成因（R45 配对 bError）/ the fault cause paired with bError
        _ePhase := E_DL_ApcPhase.eFault; // 迁故障相 / migrate to the fault phase
    ELSIF rtProbe.Q THEN // 探针触发沿：锁存位置（锁存纪律：本拍一次写入）/ the trigger edge, the position latches once this scan
        _fLatch := fPosAct; // 锁存副本写入（评价唯一来源）/ the latched copy, the only evaluation source
        _ePhase := E_DL_ApcPhase.eRetract; // 迁回退相 / migrate to the retract phase
    ELSIF tonProbe.Q THEN // 慢探超时 / the probe timed out
        _bFault := TRUE; // 置故障锁存 / raise the fault latch
        _eFaulC := E_DL_ApcFault.eNoTrigger; // 故障级成因（R45 配对 bError）/ the fault cause paired with bError
        _ePhase := E_DL_ApcPhase.eFault; // 迁故障相 / migrate to the fault phase
    END_IF

E_DL_ApcPhase.eRetract: // 回退相：退回安全距 / the retract phase, back to the safe distance
    fVelCmd := fVelFast; // 回退用快进档（反向由外部换向）/ the retract uses the fast gear, the direction is external
    IF (NOT bEnable) OR bAbort THEN // 失能或中止 / disabled or aborting
        _ePhase := E_DL_ApcPhase.eIdle; // 回空闲相 / back to idle
    ELSIF fPosAct <= (_fLatch - fBackDist) THEN // 已退到安全距 / the safe distance is reached
        _ePhase := E_DL_ApcPhase.eSettle; // 迁稳定相 / migrate to the settle phase
    ELSIF tonRetr.Q THEN // 回退超时 / the retract timed out
        _bFault := TRUE; // 置故障锁存 / raise the fault latch
        _eFaulC := E_DL_ApcFault.eNoTrigger; // 故障级成因（回退超时归并触发缺失带，R190 同带子带）/ the fault cause, the retract timeout rides the trigger band
        _ePhase := E_DL_ApcPhase.eFault; // 迁故障相 / migrate to the fault phase
    END_IF

E_DL_ApcPhase.eSettle: // 稳定相：速度归零驻留 / the settle phase, the velocity zeroes and dwells
    fVelCmd := 0.0; // 速度命令归零 / the velocity command zeroes
    IF (NOT bEnable) OR bAbort THEN // 失能或中止 / disabled or aborting
        _ePhase := E_DL_ApcPhase.eIdle; // 回空闲相 / back to idle
    ELSIF tonSettle.Q THEN // 稳定驻留窗已过 / the dwell window elapsed
        _ePhase := E_DL_ApcPhase.eRecord; // 迁记录相 / migrate to the record phase
    END_IF

E_DL_ApcPhase.eRecord: // 记录相：锁存样本入环并评价 / the record phase, the latched sample enters the ring and the verdict runs
    IF (NOT bEnable) OR bAbort THEN // 失能或中止 / disabled or aborting
        _ePhase := E_DL_ApcPhase.eIdle; // 回空闲相 / back to idle
    ELSE // 记录与评价 / the recording and the verdict
        IF _nCnt < 20 THEN // 样本环未满（钳定后重复数不超过 20）/ the ring is not full
            _nCnt := _nCnt + 1; // 样本数递增 / increment the sample count
            _anMeas[_nCnt] := _fLatch; // 锁存值入环（非实时镜像）/ the latched value enters the ring, never the live mirror
        END_IF
        IF _nCnt >= _nRepeat THEN // 样本齐 / the samples are complete
            _fMax := _anMeas[1]; // 最大值起步 / start the maximum
            _fMin := _anMeas[1]; // 最小值起步 / start the minimum
            _fSum := 0.0; // 和清零 / clear the sum
            _nI := 1; // 游标起步 / start the cursor
            _nGuard := 0; // 守护清零 / clear the guard
            WHILE (_nI <= _nCnt) AND (_nGuard < 20) DO // 时间序遍历样本环 / traverse the sample ring in time order
                _nGuard := _nGuard + 1; // 守护递增 / increment the guard
                IF _anMeas[_nI] > _fMax THEN // 最大值刷新 / refresh the maximum
                    _fMax := _anMeas[_nI]; // 更新 / update
                END_IF
                IF _anMeas[_nI] < _fMin THEN // 最小值刷新 / refresh the minimum
                    _fMin := _anMeas[_nI]; // 更新 / update
                END_IF
                _fSum := _fSum + _anMeas[_nI]; // 和累计 / accumulate the sum
                _nI := _nI + 1; // 游标递增 / increment the cursor
            END_WHILE
            IF (_fMax - _fMin) > fScatterTol THEN // 离散度超差 / the scatter is over the tolerance
                _bFault := TRUE; // 置故障锁存 / raise the fault latch
                _eFaulC := E_DL_ApcFault.eScatterHigh; // 故障级成因（R45 配对 bError）/ the fault cause paired with bError
                _ePhase := E_DL_ApcPhase.eFault; // 迁故障相 / migrate to the fault phase
            ELSE // 离散度合格，出结论 / the scatter passes, the verdict is raised
                fMeasPos := _fSum / INT_TO_LREAL(_nCnt); // 均值结论，除子已证大于零 / the mean verdict with a proven divisor
                _bDoneInt := TRUE; // 有效脉冲内部位置位（统一出口映射，R187）/ raise the internal valid bit
                _ePhase := E_DL_ApcPhase.eDone; // 迁完成相 / migrate to the done phase
            END_IF
        ELSE // 样本未齐，再来一轮 / the samples are incomplete, another round
            _ePhase := E_DL_ApcPhase.eFastApproach; // 迁快进相 / migrate to the fast approach phase
        END_IF
    END_IF

E_DL_ApcPhase.eDone: // 完成相：结论驻留，速度归零，等复位或新启动 / the done phase, the verdict holds until reset or a new start
    fVelCmd := 0.0; // 速度命令归零 / the velocity command zeroes
    IF (NOT bEnable) OR bAbort OR rtStart.Q THEN // 失能、中止或新启动沿 / disabled, aborting or a new start edge
        _ePhase := E_DL_ApcPhase.eIdle; // 回空闲相 / back to idle
    END_IF

E_DL_ApcPhase.eFault: // 故障相：速度归零，成因锁存，等复位沿 / the fault phase, the velocity zeroes until the reset edge
    fVelCmd := 0.0; // 速度安全侧归零 / the velocity takes the safe side zero
    IF NOT bEnable THEN // 失能 / disabled
        _ePhase := E_DL_ApcPhase.eIdle; // 迁未使能相 / migrate to idle
    END_IF

ELSE // 非法相位兜底（R128）/ the illegal phase fallback
    _bFault := TRUE; // 置故障锁存 / raise the fault latch
    _eFaulC := E_DL_ApcFault.ePhaseBad; // 故障级成因（R45 配对 bError）/ the fault cause paired with bError
    _ePhase := E_DL_ApcPhase.eFault; // 迁故障相 / migrate to the fault phase
END_CASE

// 段 5｜统一出口 / segment 5, the unified outlet
bMeasValid := _bDoneInt; // 有效脉冲映射本拍值 / map the valid pulse for this scan
_bDoneInt := FALSE; // 映射后立即撤销，保证单拍宽度（R187 两段式）/ revoke right after mapping
nMeasCnt := _nCnt; // 已完成测量次数出口 / the completed count outlet
IF _bFault THEN // 故障锁存优先 / the fault latch takes priority
    eFault := _eFaulC; // 故障级成因锁存回放（R152）/ the fault cause replayed from the latch
ELSE
    eFault := E_DL_ApcFault.eNone; // 无锁存即无成因 / no latch, no cause
END_IF
ePhase := _ePhase; // 相位出口单点映射 / single point phase outlet mapping
bError := _bFault; // 故障标志与锁存位同源 / the fault flag shares the latch source
END_FUNCTION_BLOCK

(* ---- FB_DL_AxisProbeTouchOffSeq.st ---- *)
(*
  FB_DL_AxisProbeTouchOffSeq —— 探针触测状态机：快进-慢进-触发记录-回退，超程与未触发超时双兜底
  分类：DL_Motion | 复杂度：3 | 轮次：R86
  开源溯源：道莅原创（clean-room 自研，纯 IEC 61131-3 通用算法），无外部代码引用
  许可证：MIT

  职责：正向（+方向）接近工件的两段式触测序列——快进到 fFastSpan 后转慢进，探针上升沿记录当前实际位置，
        随后反向回退到 fRetractDist 之外并驻留，最后给出 xDone。
  输入契约：fPosAct 为轴实际位置 [mm]（由调用方从轴接口取，本件不引用任何物理地址）；
            fFastVel / fSlowVel > 0；fSoftMax > fSoftMin；fRetractDist > 0；tTimeout / tDwell 为标准 TIME。
  输出契约：fVelCmd 速度指令 [mm/s]（快进为正、回退为负）；fProbePos 记录的触发位置 [mm]；
            xDone / xFault 均为锁存位，只在启动沿清除；eStateOut 为当前相枚举。
  边界：① 双兜底——超程（fPosAct 越 fSoftMax / fSoftMin）与未触发超时（tonTimeout.Q）均迁 FAULT；
        ② FAULT 保持最后有效 fProbePos 并置 xFault，不按当下输入重新推断；
        ③ 两个 TON 实例一律在 CASE 之外无条件每周期调用（R7）；超时定时器用锁存位单稳态自复位（R188）；
        ④ 除零防护：无除法；浮点比较一律容差 DL_EPS；⑤ 零全局耦合、零物理地址、零库件依赖。
*)

(*-----------------------------------------------------------------------------
 * 枚举: E_DL_ProbState（探针触测相，归属本文件，全库唯一定义）
 *----------------------------------------------------------------------------*)
TYPE E_DL_ProbState :
(
    eIdle       := 0,   // 空闲待启动 [—] / Idle, waiting for the start edge
    eFastApproach := 1, // 快进相（正向快速接近） [—] / Fast approach phase, positive direction
    eSlowApproach := 2, // 慢进相（正向精细接近） [—] / Slow approach phase, positive direction
    eRecord     := 3,   // 触发记录相（单拍锁存探针位置） [—] / Record phase, latches the probe position
    eRetract    := 4,   // 回退相（反向离开工件） [—] / Retract phase, negative direction
    eDwell      := 5,   // 驻留相（零速等待稳定） [—] / Dwell phase at zero velocity
    eFault      := 6    // 故障相（超程 / 超时 / 参数非法，锁存） [—] / Fault phase, latched
);
END_TYPE

FUNCTION_BLOCK FB_DL_AxisProbeTouchOffSeq
VAR_INPUT
    xEnable      : BOOL  := TRUE;   // 使能，FALSE 时任意相立即回空闲 [—] / Enable, false resets to idle from any phase
    xStart       : BOOL  := FALSE;  // 启动（上升沿开始一次触测） [—] / Start, a rising edge begins one probing cycle
    fPosAct      : LREAL := 0.0;    // 轴实际位置（由调用方传入） [mm] / The actual axis position fed by the caller
    xProbeTrig   : BOOL  := FALSE;  // 探针触发原始信号 [—] / The raw probe trigger signal
    fFastVel     : LREAL := 20.0;   // 快进速度（正值，正向） [mm/s] / Fast approach velocity, positive
    fSlowVel     : LREAL := 2.0;    // 慢进速度（正值，正向） [mm/s] / Slow approach velocity, positive
    fFastSpan    : LREAL := 50.0;   // 快进段行程（自启动位置起算） [mm] / The fast approach span from the start position
    fSoftMax     : LREAL := 200.0;  // 软限位上界 [mm] / The soft limit upper bound
    fSoftMin     : LREAL := -10.0;  // 软限位下界 [mm] / The soft limit lower bound
    fRetractDist : LREAL := 5.0;    // 回退距离（自记录位置起算） [mm] / The retract distance from the recorded position
    tTimeout     : TIME  := T#5S;   // 未触发超时门限 [s] / The not triggered timeout threshold
    tDwell       : TIME  := T#200MS;// 回退后驻留时间 [s] / The dwell time after retracting
END_VAR
VAR_OUTPUT
    fVelCmd    : LREAL;                     // 速度指令（带方向） [mm/s] / The velocity command with direction
    fProbePos  : LREAL;                     // 记录的探针触发位置 [mm] / The recorded probe trigger position
    xBusy      : BOOL;                      // 触测进行中 [—] / Probing in progress
    xDone      : BOOL;                      // 序列完成（锁存，启动沿清除） [—] / Sequence done, latched and cleared by the start edge
    xFault     : BOOL;                      // 故障（锁存，启动沿清除） [—] / Fault, latched and cleared by the start edge
    eStateOut  : E_DL_ProbState;            // 当前相枚举 [—] / The current phase enumeration
END_VAR
VAR
    eState        : E_DL_ProbState;         // 内部相（与 eStateOut 同步发布） [—] / Internal phase mirrored to eStateOut
    xStartPrev    : BOOL;                   // 启动信号上拍快照 [—] / Previous scan snapshot of xStart
    xProbePrev    : BOOL;                   // 探针信号上拍快照 [—] / Previous scan snapshot of xProbeTrig
    xStartEdge    : BOOL;                   // 本拍启动上升沿 [—] / The start rising edge this scan
    xProbeEdge    : BOOL;                   // 本拍探针上升沿 [—] / The probe rising edge this scan
    xTimeoutLatch : BOOL;                   // 超时锁存位（单稳态自复位用） [—] / The timeout latch used for the monostable reset
    xApproaching  : BOOL;                   // 处于接近两相（超时定时器使能条件） [—] / In an approach phase, the timer enable
    xParamBad     : BOOL;                   // 参数非法标志 [—] / Parameter invalid flag
    fPosRef       : LREAL;                  // 启动时的位置基准 [mm] / The position reference captured at the start edge
    fProbeLast    : LREAL;                  // 最后有效触发位置 [mm] / The last valid trigger position
    tonTimeout    : TON;                    // 未触发超时定时器（CASE 外无条件调用） [—] / The not triggered timeout timer
    tonDwell      : TON;                    // 回退后驻留定时器（CASE 外无条件调用） [—] / The dwell timer after retracting
END_VAR
VAR CONSTANT
    DL_EPS  : LREAL := 1.0E-9;              // 浮点比较容差 [—] / The floating point comparison tolerance
    DL_ZERO : LREAL := 0.0;                 // 浮点零常量 [—] / The floating point zero constant
END_VAR

// 段 1｜周期无条件刷新：沿提取、使能判定、出口指令预置
xStartEdge := xStart AND NOT xStartPrev;                  // 启动上升沿提取 / extract the start rising edge
xProbeEdge := xProbeTrig AND NOT xProbePrev;              // 探针上升沿提取 / extract the probe rising edge
xApproaching := (eState = E_DL_ProbState.eFastApproach) OR (eState = E_DL_ProbState.eSlowApproach); // 接近两相判定
xBusy := FALSE;                                           // 忙碌位预置假，接近 / 回退 / 驻留相置真 / preset busy false
fVelCmd := DL_ZERO;                                       // 速度指令预置零，各相按需置值 / preset the velocity command zero

// 段 2｜两个定时器无条件调用（R7：不在 IF / CASE 内调用）
tonTimeout(IN := xApproaching AND NOT xTimeoutLatch, PT := tTimeout); // 未触发超时：接近相且未锁存时计时
tonDwell(IN := (eState = E_DL_ProbState.eDwell) AND NOT tonDwell.Q, PT := tDwell); // 驻留：驻留相计时，Q 到后自复位
IF tonTimeout.Q THEN                                      // 超时到（首次到达即锁存） / the timeout elapsed
    xTimeoutLatch := TRUE;                                // 锁存超时位，复位定时器 IN / latch so the timer resets
END_IF

// 段 2.5｜使能总闸（R86 审校 BLOCK 修复）：撤使能须从任意运动相立即停机，不能只在空闲相判
IF (NOT xEnable) AND (eState <> E_DL_ProbState.eFault) THEN   // 撤使能且当前非故障相 / enable dropped while not faulted
    eState := E_DL_ProbState.eIdle;                           // 强制回空闲相 / force the state back to idle
    fVelCmd := DL_ZERO;                                       // 速度指令立即清零，禁止带着速度指令穿越 / zero the velocity command at once
    xBusy := FALSE;                                           // 清忙碌位 / clear the busy flag
END_IF

// 段 3｜主状态机（ENUM + CASE，ELSE 拦截非法相）
CASE eState OF

    E_DL_ProbState.eIdle:
        IF NOT xEnable THEN                               // 未使能时保持空闲并清锁存 / stay idle and clear the latches
            xDone := FALSE;                               // 清完成锁存 [—] / clear the done latch
            xFault := FALSE;                              // 清故障锁存 [—] / clear the fault latch
            xTimeoutLatch := FALSE;                       // 清超时锁存 [—] / clear the timeout latch
        END_IF
        IF xStartEdge AND xEnable THEN                    // 使能下的启动沿 / a start edge while enabled
            xDone := FALSE;                               // 启动沿清完成锁存 [—] / clear the done latch on the start edge
            xFault := FALSE;                              // 启动沿清故障锁存 [—] / clear the fault latch on the start edge
            xTimeoutLatch := FALSE;                       // 启动沿清超时锁存 [—] / clear the timeout latch on the start edge
            xParamBad := FALSE;                           // 参数闸标志复位 / reset the parameter gate flag
            IF fFastVel <= DL_ZERO THEN                   // 快进速度非正 / the fast velocity is non positive
                xParamBad := TRUE;                        // 判参数非法 / mark the parameters invalid
            END_IF
            IF fSlowVel <= DL_ZERO THEN                   // 慢进速度非正 / the slow velocity is non positive
                xParamBad := TRUE;                        // 判参数非法 / mark the parameters invalid
            END_IF
            IF fFastSpan < DL_ZERO THEN                   // 快进行程为负 / the fast span is negative
                xParamBad := TRUE;                        // 判参数非法 / mark the parameters invalid
            END_IF
            IF fRetractDist <= DL_ZERO THEN               // 回退距离非正 / the retract distance is non positive
                xParamBad := TRUE;                        // 判参数非法 / mark the parameters invalid
            END_IF
            IF fSoftMax <= fSoftMin THEN                  // 软限位上下界倒置 / the soft limits are inverted
                xParamBad := TRUE;                        // 判参数非法 / mark the parameters invalid
            END_IF
            IF (fPosAct > fSoftMax) OR (fPosAct < fSoftMin) THEN // 起始位置已在限位外 / already outside the soft limits
                xParamBad := TRUE;                        // 判参数非法 / mark the parameters invalid
            END_IF
            IF xParamBad THEN                             // 任一闸判失败 / any gate failed
                eState := E_DL_ProbState.eFault;          // 迁入故障相 / enter the fault phase
                xFault := TRUE;                           // 置故障锁存 [—] / raise the fault latch
            ELSE
                fPosRef := fPosAct;                       // 捕获启动位置基准 [mm] / capture the start position reference
                fProbeLast := fPosAct;                    // 触发位置初值取启动位置 [mm] / the initial trigger position
                fProbePos := fProbeLast;                  // 出口同步初值 [mm] / mirror the outlet value
                eState := E_DL_ProbState.eFastApproach;   // 迁入快进相 / enter the fast approach phase
            END_IF
        END_IF

    E_DL_ProbState.eFastApproach:
        fVelCmd := fFastVel;                              // 快进速度指令 [mm/s] / the fast approach velocity command
        xBusy := TRUE;                                    // 置忙碌位 [—] / raise the busy flag
        IF xProbeEdge THEN                                // 探针已触发 / the probe already triggered
            eState := E_DL_ProbState.eRecord;             // 直接进入记录相（本拍合法事件优先） / go straight to record
        ELSIF (fPosAct > fSoftMax) OR (fPosAct < fSoftMin) THEN // 软限位超程（兜底一） / the soft limit is exceeded
            eState := E_DL_ProbState.eFault;              // 迁入故障相 / enter the fault phase
            xFault := TRUE;                               // 置故障锁存 [—] / raise the fault latch
            fVelCmd := DL_ZERO;                           // 故障即切零速 [mm/s] / cut the velocity to zero
        ELSIF (fPosAct - fPosRef) >= fFastSpan THEN       // 快进行程走满 / the fast span is used up
            eState := E_DL_ProbState.eSlowApproach;       // 转入慢进相 / switch to the slow approach phase
        ELSIF xTimeoutLatch THEN                          // 未触发超时（兜底二） / the not triggered timeout fired
            eState := E_DL_ProbState.eFault;              // 迁入故障相 / enter the fault phase
            xFault := TRUE;                               // 置故障锁存 [—] / raise the fault latch
            fVelCmd := DL_ZERO;                           // 故障即切零速 [mm/s] / cut the velocity to zero
        END_IF

    E_DL_ProbState.eSlowApproach:
        fVelCmd := fSlowVel;                              // 慢进速度指令 [mm/s] / the slow approach velocity command
        xBusy := TRUE;                                    // 置忙碌位 [—] / raise the busy flag
        IF xProbeEdge THEN                                // 探针触发 / the probe triggered
            eState := E_DL_ProbState.eRecord;             // 进入记录相（本拍合法事件优先） / enter the record phase first
        ELSIF (fPosAct > fSoftMax) OR (fPosAct < fSoftMin) THEN // 软限位超程（兜底一） / the soft limit is exceeded
            eState := E_DL_ProbState.eFault;              // 迁入故障相 / enter the fault phase
            xFault := TRUE;                               // 置故障锁存 [—] / raise the fault latch
            fVelCmd := DL_ZERO;                           // 故障即切零速 [mm/s] / cut the velocity to zero
        ELSIF xTimeoutLatch THEN                          // 未触发超时（兜底二） / the not triggered timeout fired
            eState := E_DL_ProbState.eFault;              // 迁入故障相 / enter the fault phase
            xFault := TRUE;                               // 置故障锁存 [—] / raise the fault latch
            fVelCmd := DL_ZERO;                           // 故障即切零速 [mm/s] / cut the velocity to zero
        END_IF

    E_DL_ProbState.eRecord:
        fProbeLast := fPosAct;                            // 锁存本次触发位置 [mm] / latch the trigger position of this cycle
        fProbePos := fProbeLast;                          // 发布到出口 [mm] / publish it to the outlet
        xBusy := TRUE;                                    // 记录拍仍算忙碌 [—] / the record scan still counts as busy
        eState := E_DL_ProbState.eRetract;                // 下一拍进入回退相 / move to the retract phase next scan
        IF fProbeLast > fSoftMax THEN                     // 记录位置越上限的不可能态兜底 / a defensive check on the record
            eState := E_DL_ProbState.eFault;              // 迁入故障相 / enter the fault phase
            xFault := TRUE;                               // 置故障锁存 [—] / raise the fault latch
        END_IF

    E_DL_ProbState.eRetract:
        fVelCmd := -fSlowVel;                             // 反向回退速度指令 [mm/s] / the negative retract velocity command
        xBusy := TRUE;                                    // 置忙碌位 [—] / raise the busy flag
        IF (fProbeLast - fPosAct) >= fRetractDist THEN    // 回退距离走满 / the retract distance is covered
            eState := E_DL_ProbState.eDwell;              // 转入驻留相 / switch to the dwell phase
            fVelCmd := DL_ZERO;                           // 驻留相速度归零 [mm/s] / zero velocity in the dwell phase
        ELSIF fPosAct < fSoftMin THEN                     // 回退越下软限位 / the lower soft limit is exceeded while retracting
            eState := E_DL_ProbState.eFault;              // 迁入故障相 / enter the fault phase
            xFault := TRUE;                               // 置故障锁存 [—] / raise the fault latch
            fVelCmd := DL_ZERO;                           // 故障即切零速 [mm/s] / cut the velocity to zero
        END_IF

    E_DL_ProbState.eDwell:
        fVelCmd := DL_ZERO;                               // 驻留相零速保持 [mm/s] / hold zero velocity during the dwell
        xBusy := TRUE;                                    // 置忙碌位 [—] / raise the busy flag
        IF tonDwell.Q THEN                                // 驻留计时到 / the dwell elapsed
            eState := E_DL_ProbState.eIdle;               // 回空闲相 / back to idle
            xDone := TRUE;                                // 置完成锁存 [—] / raise the done latch
        END_IF

    E_DL_ProbState.eFault:
        fVelCmd := DL_ZERO;                               // 故障相速度指令归零 [mm/s] / the fault phase velocity is zero
        fProbePos := fProbeLast;                          // 故障相保持最后有效触发位置 [mm] / hold the last valid trigger position
        xFault := TRUE;                                   // 故障锁存回放 [—] / replay the latched fault flag
        IF (NOT xStart) AND NOT xEnable THEN              // 撤启动且撤使能 / start released and enable dropped
            eState := E_DL_ProbState.eIdle;               // 唯一解除路径：该条件沿回空闲 / the only clear edge back to idle
            xTimeoutLatch := FALSE;                       // 同时清超时锁存 [—] / clear the timeout latch as well
        END_IF

ELSE
    eState := E_DL_ProbState.eFault;                      // 非法枚举值一律拦入故障相 / trap any illegal phase value
    xFault := TRUE;                                       // 置故障锁存 [—] / raise the fault latch
    fVelCmd := DL_ZERO;                                   // 速度指令归零 [mm/s] / the velocity command is zero
    fProbePos := fProbeLast;                              // 保持最后有效触发位置 [mm] / hold the last valid trigger position
END_CASE

// 段 4｜相枚举出口发布 + 输入上拍快照（主体末尾，保证本拍沿检测用上拍值）
eStateOut := eState;                                      // 相枚举统一出口（单点发布） / the single point phase outlet
xStartPrev := xStart;                                     // 刷新启动上拍快照 / refresh the start snapshot
xProbePrev := xProbeTrig;                                 // 刷新探针上拍快照 / refresh the probe snapshot
END_FUNCTION_BLOCK

(* ---- FB_DL_AxisRelativeMove.st ---- *)
(*==============================================================================
 * 组件名称 (Component)  : FB_DL_AxisRelativeMove
 * 所属子库 (Sublibrary) : DL_Motion
 * 当前版本 (Version)    : 1.0.0
 * 组件分类 (Category)   : 功能块（FUNCTION_BLOCK）· 单轴相对定位与链式步进封装 · 工艺上层件
 * 兼容性   (Platform)   : CODESYS 3.5 / TwinCAT 3 / 汇川 InoProShop / Schneider
 *                         Machine Expert；仅依赖 Standard.library（R_TRIG / MIN /
 *                         MAX / ABS），零厂商方言
 * 接口依赖 (Depends)    : I_DL_MotionAxis / E_DL_AxisState（既有契约，Round 05）
 * 功能描述 (Function)   : 单轴相对定位（MC_MoveRelative 语义）与连续累加步进
 *                         控制封装。经轴接口引用驱动轴体：上升沿发起
 *                         MoveRelative，轮询轴状态回待机判步完成；链式模式下
 *                         到位后自动连续执行下一步，步间距即 fDistance，上层
 *                         运行中递增 nChainTarget 即实现无上限累加步进。
 * 设计要点 (Key notes)  : ① 启动门禁：仅在轴待机态发起；fVel/fAcc 非正值或
 *                           非有限值 → 拒绝启动并置信息级 0004_0106（与
 *                           FB_DL_AxisHomingSeq 同码同义：参数门禁拒绝，共用
 *                           留档）；
 *                         ② 指令被轴拒绝（返回 FALSE）→ 0004_0220 故障级
 *                           锁存；bAbort 或轴故障 → 受控 Stop + 0004_0221
 *                           故障级锁存；两锁存码仅新执行沿解除（R15：锁存型
 *                           故障只在解除路径清码）；
 *                         ③ 链式步进：步完成后隔一拍自动再发（轴待机确认后
 *                           消费），bDone 每步置位保持至下一步启动；
 *                         ④ 本块为事件型 + 轮询状态组件，免首扫（R23），无
 *                           连续量同步语义，不设初始化跟踪逻辑。
 * 开源溯源 (Origin)     : 原创实现（参考 PLCopen Part 1-6 MC_MoveRelative 公开
 *                         语义与西门子 Motion Control 对象语义，clean-room）。
 *                         仅提取公开指令动词与参数域；实现与命名 100% 自有，
 *                         未参考任何厂商源码行。
 * 验收向量 (Acceptance) :
 *   V1 单步链：执行沿→MoveRelative 受理→轮询回待机→bDone+计数+1；
 *   V2 链式 3 步：bChainMode+target=3 → 连续 3 步逐拍推进，bChainDone 置位；
 *   V3 目标递增累加：运行中 nChainTarget 3→5 → 链不中断续跑第 4、5 步；
 *   V4 指令被拒：轴非待机态受理失败 → 0004_0220 锁存，新执行沿解除；
 *   V5 中止：运行中 bAbort → 受控 Stop + 0004_0221；
 *   V6 状态门禁：轴故障态执行沿 → 拒绝并置信息级 0004_0106，轴状态不变。
 * 故障码表 (Error codes):
 *   16#0004_0106【信息级】启动门禁/参数门禁拒绝（与 FB_DL_AxisHomingSeq 同码
 *   同义，共用留档）；16#0004_0220【故障级】定位指令被轴拒绝（锁存）；
 *   16#0004_0221【故障级】中止/轴故障中断（锁存）；16#0004_0201【故障级】
 *   非法状态兜底（沿用族码，与 FB_DL_SingleAxis 同码同义，复用留档）。
 * 修订历史 (Revision)   :
 *   2026-11-15  v1.0.0  首版入库（Round 06 · DL_Motion 回零/运动族）
 *   2026-11-15  v1.0.1  R11 修复：枚举成员分隔符笔误，eMoving 行误写单冒号 `:`（枚举成员赋值须用 `:=`），三平台编译阻断已消除，数值与语义不变。
 *                       R11 fix: enum member separator erratum, `:` -> `:=` on one member.
 *============================================================================*)

(*-----------------------------------------------------------------------------
 * 调用示例 (Instance guide)：
 *   fbRel.iAxis := fbAxis;                        // 接口依赖注入
 *   fbRel(bCmdExecute := bDoStep, fDistance := 25.0, // 周期调用
 *         fVel := 100.0, fAcc := 1000.0,
 *         bChainMode := TRUE, nChainTarget := 10);
 *   连续累加步进：运行中每检测到一件料即 nChainTarget := nChainTarget + 1，
 *   链式机制自动续跑，无需停止重启链。
 *----------------------------------------------------------------------------*)

(*-----------------------------------------------------------------------------
 * 常见误用与现场提示 (Field notes)：
 *   1 本块仅在轴待机态发起定位，轴受控停止中/故障态一律拒绝；中止后轴自行
 *     减速回待机，无需上层等待即可发新执行沿。
 *   2 uStepsDone 在每次执行沿清零重新计数；跨链累计请上层自行汇总。
 *   3 bAbort 电平生效：运行中置 TRUE 立即受控停车并锁存 0004_0221，撤除
 *     不自动恢复运行；重新执行需新的 bCmdExecute 上升沿。
 *----------------------------------------------------------------------------*)

(*-----------------------------------------------------------------------------
 * 枚举: E_DL_RelStep（归属 DL_Motion，与 FB_DL_AxisRelativeMove 同文件）
 * 含义: 相对定位内部步进枚举（本块私有配套，外部仅作诊断参考）。
 *----------------------------------------------------------------------------*)
{attribute 'strict'}
{attribute 'qualified_only'}
TYPE E_DL_RelStep :
(
    eIdle   := 0,    // 空闲：等待执行沿 / Idle: waiting for execute edge
    eMoving := 10    // 定位进行中：轮询轴状态回待机 / Moving: polling axis back to standstill
) UINT;
END_TYPE

FUNCTION_BLOCK FB_DL_AxisRelativeMove
VAR_INPUT
    bCmdExecute   : BOOL := FALSE;      // 执行指令（Execute command），上升沿生效
    fDistance     : REAL := 0.0;        // 相对位移（Relative distance）[mm]，带符号，负值=负向
    fVel          : REAL := 100.0;      // 运行速度（Run velocity）[mm/s]，正值，默认 100.0
    fAcc          : REAL := 1000.0;     // 加减速度（Acceleration）[mm/s²]，正值，默认 1000.0
    bChainMode    : BOOL := FALSE;      // 链式步进模式（Chain mode），TRUE=到位后自动连续执行下一步
    nChainTarget  : UDINT := 1;         // 链式目标步数（Chain target steps），0=按 1 步处理；运行中递增即累加步进
    bAbort        : BOOL := FALSE;      // 中止（Abort），电平生效 → 轴受控停止
END_VAR
VAR_IN_OUT
    iAxis         : I_DL_MotionAxis;    // 轴接口引用（Axis reference），由上层注入实现块实例
END_VAR
VAR_OUTPUT
    bBusy         : BOOL := FALSE;      // 定位进行中（Move busy）
    bDone         : BOOL := FALSE;      // 单步完成（Step done），每步置位保持至下一步启动
    bChainDone    : BOOL := FALSE;      // 链式目标完成（Chain target reached）
    uStepsDone    : UDINT := 0;         // 本次链累计完成步数（Steps done），执行沿清零
    uErrorId      : UDINT := 0;         // 末次事件码（Last error code），段位 16#0004_xxxx
END_VAR
VAR
    eStep         : E_DL_RelStep := E_DL_RelStep.eIdle; // 内部步进状态（Internal step state）
    bFaultLatch   : BOOL := FALSE;      // 故障锁存标志（Fault latch），0004_0220/0221 锁存载体
    bParamOk      : BOOL := FALSE;      // 参数门禁通过标志（Parameter gate pass flag），逐拍重算
    bWaitNext     : BOOL := FALSE;      // 链式步间一拍间隔标志（Inter-step one-scan wait flag）
    bAbortDone    : BOOL := FALSE;      // 中止停止指令已发标志（Abort stop issued flag），单发化
    uChainTgt     : UDINT := 1;         // 生效链式目标（Effective chain target），下限钳位 1
    fVelEff       : REAL := 100.0;      // 生效运行速度（Effective velocity）[mm/s]，防除零兜底
    fAccEff       : REAL := 1000.0;     // 生效加减速度（Effective acceleration）[mm/s²]，防除零兜底
    rtrigExec     : R_TRIG;             // 执行指令上升沿（Rising edge of execute command）
END_VAR
VAR CONSTANT
    DL_REL_INF_MAX   : REAL := 1.0E30;  // 有限值判定幅值上限（Finite-value magnitude bound）[mm 或 mm/s]
    DL_REL_EPS       : REAL := 1.0E-6;  // 浮点判零容差（Float zero tolerance）
    DL_REL_PAR_FLOOR : REAL := 1.0E-3;  // 速度/加速度参数下限（Velocity and acceleration floor）[mm/s 或 mm/s²]
END_VAR

METHOD IssueMove : BOOL
VAR_INPUT
END_VAR
IssueMove := iAxis.MoveRelative(fDistance, fVelEff, fAccEff);  // 转发轴接口，受理结果即返回值
    END_METHOD

// 段 1｜沿检测无条件周期刷新（R7 红线，严禁置于分支内）
rtrigExec(CLK := bCmdExecute);

// 段 2｜接口引用有效性防御：未注入轴引用则清输出退出（不产生误动作）
IF iAxis = 0 THEN
    bBusy := FALSE;
    RETURN;
END_IF

// 段 3｜参数门禁逐拍重算（公约 0.8）：非法仅封锁启动，运行中不中断
bParamOk := (fDistance = fDistance) AND (fVel = fVel) AND (fAcc = fAcc)
        AND (ABS(fDistance) <= DL_REL_INF_MAX) AND (fVel <= DL_REL_INF_MAX)
        AND (fAcc <= DL_REL_INF_MAX)
        AND (fVel > DL_REL_PAR_FLOOR) AND (fAcc > DL_REL_PAR_FLOOR);
fVelEff := MAX(fVel, DL_REL_PAR_FLOOR);          // 生效速度下限兜底 [mm/s]，防除零
fAccEff := MAX(fAcc, DL_REL_PAR_FLOOR);          // 生效加速度下限兜底 [mm/s²]，防除零

// 段 4｜事件码管理（R15）：瞬时码逐拍重算，锁存码仅在解除路径（新执行沿）清
IF NOT bFaultLatch THEN
    uErrorId := 0;
END_IF

// 段 5｜定位状态机（ENUM + CASE + ELSE 兜底）
CASE eStep OF

    E_DL_RelStep.eIdle:                          // 空闲态：等待执行沿与门禁
        bBusy := FALSE;
        IF rtrigExec.Q THEN
            bFaultLatch := FALSE;                // 新执行沿：锁存码解除路径（R15）
            IF NOT bParamOk THEN
                uErrorId := 16#0004_0106;        // 参数门禁拒绝（信息级）
            ELSIF iAxis.eState <> E_DL_AxisState.eStandstill THEN
                uErrorId := 16#0004_0106;        // 轴非待机态，拒绝发起（信息级）
            ELSE
                uChainTgt := 1;                  // 非链式恒为单步目标 [步]
                IF bChainMode THEN uChainTgt := MAX(nChainTarget, 1); END_IF  // 链式目标下限钳位 1
                uStepsDone := 0;                 // 本次链计数清零
                bDone := FALSE;
                bChainDone := FALSE;
                bWaitNext := FALSE;
                bAbortDone := FALSE;
                IF IssueMove() THEN
                    eStep := E_DL_RelStep.eMoving;
                    bBusy := TRUE;
                ELSE
                    bFaultLatch := TRUE;         // 指令被轴拒绝：故障级锁存
                    uErrorId := 16#0004_0220;
                END_IF
            END_IF
        END_IF

    E_DL_RelStep.eMoving:                        // 定位态：轮询轴状态，链式自动续步
        bBusy := TRUE;
        IF bAbort OR iAxis.bError THEN
            IF NOT bAbortDone THEN
                iAxis.Stop();                    // 中止/轴故障：受控停车单发
                bAbortDone := TRUE;
            END_IF
            bFaultLatch := TRUE;                 // 故障级锁存（R15：仅新执行沿解除）
            uErrorId := 16#0004_0221;
            bBusy := FALSE;
            eStep := E_DL_RelStep.eIdle;
        ELSIF bWaitNext THEN
            bWaitNext := FALSE;                  // 链式步间隔拍：下一拍自动再发（连续累加步进语义）
            IF NOT IssueMove() THEN
                bFaultLatch := TRUE;             // 续步指令被拒：故障级锁存
                uErrorId := 16#0004_0220;
                bBusy := FALSE;
                eStep := E_DL_RelStep.eIdle;
            END_IF
        ELSIF iAxis.eState = E_DL_AxisState.eStandstill THEN
            bDone := TRUE;                       // 单步完成：置位保持至下一步启动
            uStepsDone := uStepsDone + 1;        // 步计数递增 [步]
            IF bChainMode AND (uStepsDone < uChainTgt) THEN
                bWaitNext := TRUE;               // 链未达目标：下一拍续步
            ELSE
                IF bChainMode THEN
                    bChainDone := TRUE;          // 链式目标完成
                END_IF
                bBusy := FALSE;
                eStep := E_DL_RelStep.eIdle;
            END_IF
        END_IF

    ELSE
        // 非法状态兜底（故障级，沿用族码 0004_0201，复用留档）
        uErrorId := 16#0004_0201;
        bFaultLatch := TRUE;
        bBusy := FALSE;
        eStep := E_DL_RelStep.eIdle;

END_CASE

(*-----------------------------------------------------------------------------
 * 方法实现（METHOD）：相对定位指令派发子过程，非阻塞，直接转发轴接口受理
 * 结果；步间距取当前 fDistance 输入值，链式运行中改位移即改步距。
 *-----------------------------------------------------------------------------*)

END_FUNCTION_BLOCK

(* ---- FB_DL_AxisRotaryShortPath.st ---- *)
(*==============================================================================
 * 组件名称 (Component)  : FB_DL_AxisRotaryShortPath
 * 所属子库 (Sublibrary) : DL_Motion
 * 当前版本 (Version)    : 1.0.0
 * 兼容性   (Platform)   : CODESYS 3.5+ / TwinCAT 3 / 汇川 InoProShop / 施耐德 Machine Expert
 *                         仅依赖 Standard.library（R_TRIG / ABS / TRUNC），零厂商私有库
 * 功能描述 (Function)   : 旋转轴（可多圈）最短路径规划。把当前任意圈数域位置归一化到 [0,360)，
 *                         再据目标角求最小转角 d：d > 180° 走反向、d < −180° 走正向；
 *                         加圈后得到绝对目标位 fTargetAbs 与圈号 nTurnIndex，并按软限做二次
 *                         校核（首选圈越限时尝试另一圈，仍越限则拒绝并置码）。
 * 角度约定 (Corner)     : **d 恰好等于 ±180° 时**：按「正方向（CW，角度增大）优先」确定为 +180°，
 *                         且 bCwOnly 为真时无论 d 正负一律转成正向等价角〔即取 +360 方向的长路径〕。
 *                         该约定写死在此处与实现一致，不得留空由调用方猜测。
 * 接口     (Interface)  : 输入 fPosAct 当前位置（可为任意圈数）、fTargetDeg 目标角（0~360）、
 *                         fSoftLoDeg / fSoftHiDeg 圈域软限、bCwOnly 单向（只允许正向）模式、
 *                         bExecute 规划触发沿、bReset 复位；输出 bShortestCw 转向建议（TRUE=正向）、
 *                         fTargetAbs 加圈后绝对目标位、nTurnIndex 目标圈号、bValid 规划有效、
 *                         eState / eCause / bError / nErrId。
 * 边界     (Boundary)   : ① 归一化一律**条件加减**，禁 MOD（负数取余在三平台不一致，R10/R48 铁律），
 *                         循环带守卫计数器，超限即置码跳出（不死循环）；
 *                         ② 圈号用 DINT 承载并带守卫上限，越界前置判，绝不静默回绕；
 *                         ③ 组态闸：fSoftHiDeg <= fSoftLoDeg、fTargetDeg 越 [0,360]、任一时恒为
 *                         NaN → 故障锁存（每个参与判据的引脚都在闸内，R151）；
 *                         ④ **整数进位点两向量已推**（R149 终审两式 2）：
 *                         向量 A：fPosAct = 720.0、fTargetDeg = 0.0 → 归一 0.0、d = 0.0，
 *                                 fTargetAbs = 720.0、nTurnIndex = 2（整除点不跳圈，不得出 1 或 3）；
 *                         向量 B：fSoftLoDeg = 0.0、fSoftHiDeg = 359.0、fTargetDeg = 360.0
 *                                 → 候选位 360.0 越上限，须尝试另一圈（0.0）并成功，**不得回绕后
 *                                 仍报越限**；
 *                         ⑤ R_TRIG 两枚（执行/复位）段 0 无条件刷新；
 *                         ⑥ 故障相迁出唯一路径 = bReset 上升沿；⑦ 零全局耦合（无 GVL / 无物理地址）。
 * 解除式   (Release)    : bReset 上升沿 ∧ 组态合法 ∧ 目标域合法 ∧ 〔当拍已求得软限内解 ∨
 *                         目标角本身落在软限区间内〕（两分支均全当拍量，R240 范式）。
 *                         自证可满足（终审两式 1）：分支 2 只依赖 fTargetDeg 与软限的当拍比较，
 *                         不依赖执行沿（若只保留依赖 _bSolved 的分支 1，未按执行时该项恒假 →
 *                         故障永久不可恢复，属 R152 恒假组合反例），故实现为双分支析取式。
 * 码表     (Codes)      : 16#0004_03B8 故障级：旋转最短路径故障总码（组态非法 / 目标角越域 /
 *                         归一化超迭代守卫 / 软限无解 / 非法相位），锁存至 bReset 上升沿，
 *                         归因由 eCause 承载（R190 单件单总码）；
 *                         16#0004_04B8 信息级：规划成功（给出转向建议与绝对目标位）。
 *                         加码反证（R90）：规划成功与「未执行」在 fTargetAbs 上可能同值（d = 0 时
 *                         目标位等于当前位置），bValid 又只是布尔位不进台账，故立一码留痕。
 *                         码段说明：0004 段故障子带 03xx / 信息子带 04xx，本件取 03B8 / 04B8
 *                         （源码实扫该两槽为空，续接同子带已用最大值，未回填碎片孔洞）。
 * 开源溯源 (Origin)     : 道莅自研 clean-room（参考旋转轴最短路径与角度归约公开算法，
 *                         零代码行复制；t1-6-plcopen 族）
 * 修订历史 (Revision)   : 2026-11-19  v1.0.0  R45 首版（批次 3 · 序号 14）
 *==============================================================================*)

TYPE E_DL_RspState :
(
    eIdle  := 0,     // 待规划触发 / Idle, awaiting execute edge
    eRun   := 10,    // 规划结果就绪 / Plan ready
    eFault := 90     // 故障锁存相 / Fault latched phase
);
END_TYPE

TYPE E_DL_RspCause :
(
    eNone       := 0,   // 无故障成因 / No cause
    eCfgIllegal := 1,   // 组态非法（软限倒置或 NaN） / Illegal configuration
    eTargetBad  := 2,   // 目标角越 [0,360] / Target angle out of domain
    eIterGuard  := 3,   // 归一化超迭代守卫 / Normalisation iteration guard tripped
    eSoftLimit  := 4,   // 软限无解（两圈均越限） / No solution inside soft limits
    eTurnGuard  := 5,   // 圈号超守卫上限 / Turn index guard tripped
    ePhaseBad   := 6    // 非法相位兜底 / Illegal phase fallback
);
END_TYPE

FUNCTION_BLOCK FB_DL_AxisRotaryShortPath
VAR_INPUT
    fPosAct     : REAL := 0.0;          // 当前位置（任意圈数域，度） [deg] / Current position in any turn domain [deg]
    fTargetDeg  : REAL := 0.0;          // 目标角，有效域 0.0 ~ 360.0 [deg] / Target angle, domain 0.0..360.0 [deg]
    fSoftLoDeg  : REAL := 0.0;          // 圈域软限下限，域 < fSoftHiDeg [deg] / Turn-domain soft limit lower bound [deg]
    fSoftHiDeg  : REAL := 1080.0;       // 圈域软限上限，域 > fSoftLoDeg [deg] / Turn-domain soft limit upper bound [deg]
    bCwOnly     : BOOL := FALSE;        // 单向模式（只允许正方向 CW） [-] / CW-only mode
    bExecute    : BOOL := FALSE;        // 规划触发，上升沿受理一次 [-] / Plan trigger, rising edge accepts once
    bReset      : BOOL := FALSE;        // 复位命令，上升沿清故障 [-] / Reset command, rising edge clears fault
END_VAR
VAR_OUTPUT
    bShortestCw : BOOL;                 // 转向建议：TRUE = 正方向（CW，角度增大） [-] / Direction advice, TRUE means CW
    fTargetAbs  : REAL;                 // 加圈后的绝对目标位 [deg] / Absolute target after turn selection [deg]
    nTurnIndex  : DINT;                 // 目标圈号（DINT 钳位承载） [圈] / Target turn index carried in DINT [turn]
    bValid      : BOOL;                 // 规划结果有效 [-] / Plan valid
    eState      : E_DL_RspState;        // 状态出口，段 6 单点映射 / State outlet
    eCause      : E_DL_RspCause;        // 故障成因出口（R190 归因唯一） / Fault cause outlet
    bError      : BOOL;                 // 故障锁存标志 [-] / Fault latch flag
    nErrId      : UDINT;                // 事件码，0 = 无事件 / Event code, 0 = no event
END_VAR
VAR
    _eState     : E_DL_RspState := E_DL_RspState.eIdle;    // 内部相位（CASE 唯一写入目标） / Internal phase
    _eCause     : E_DL_RspCause := E_DL_RspCause.eNone;    // 故障成因锁存（锁存量） / Latched cause
    rtExec      : R_TRIG;               // 执行沿实例，段 0 无条件调用 / Execute edge
    rtReset     : R_TRIG;               // 复位沿实例，段 0 无条件调用 / Reset edge
    _fNorm      : REAL;                 // 归一化角（[0,360) 当拍量） [deg] / Normalised angle this scan [deg]
    _fDiff      : REAL;                 // 最小转角候选（当拍量） [deg] / Candidate shortest angle [deg]
    _fAbsCand   : REAL;                 // 候选绝对目标位（当拍量） [deg] / Candidate absolute target [deg]
    _fTmp       : REAL;                 // 圈号求解临时量（当拍量） [deg] / Temporary value for turn index
    _nIter      : DINT;                 // 归一化迭代计数（当拍量） [次] / Normalisation iteration count
    _nTurnCalc  : DINT;                 // 圈号求解值（当拍量） [圈] / Turn index solving value
    _bNonFin    : BOOL;                 // 输入非有限当拍量 [-] / Non-finite input this scan
    _bCfgBad    : BOOL;                 // 组态非法当拍量 [-] / Illegal configuration
    _bTargetBad : BOOL;                 // 目标角越域当拍量 [-] / Target out of domain
    _bIterBad   : BOOL;                 // 迭代守卫触发当拍量 [-] / Iteration guard tripped
    _bTurnBad   : BOOL;                 // 圈号守卫触发当拍量 [-] / Turn guard tripped
    _bSolved    : BOOL;                 // 软限求解成功当拍量 [-] / Solved inside soft limits
    _bFault     : BOOL;                 // 故障锁存位（锁存量） / Latched fault bit
    _uFault     : UDINT;                // 故障码锁存（锁存量） / Latched fault code
    _uInfo      : UDINT;                // 信息码，每拍重算 / Info code, recomputed each scan
END_VAR
VAR CONSTANT
    DL_FLOAT_EPS : REAL := 1.0E-4;      // 角度判等容差（度级精度） [deg] / Angle epsilon at degree resolution [deg]
    DL_FULL_TURN : REAL := 360.0;       // 整圈角度，编译期常量 [deg] / Full turn constant [deg]
    DL_HALF_TURN : REAL := 180.0;       // 半圈角度，编译期常量 [deg] / Half turn constant [deg]
    DL_ITER_MAX  : DINT := 1000;        // 归一化迭代守卫上限 [次] / Normalisation iteration guard [count]
    DL_TURN_MAX  : DINT := 100000;      // 圈号守卫绝对值上限 [圈] / Turn index absolute guard [turn]
END_VAR

(* —— 段 0：当拍量派生 + 沿实例无条件周期刷新 —— *)
_bNonFin := (fPosAct <> fPosAct) OR (fTargetDeg <> fTargetDeg)                            // NaN 自反判（判等禁令唯一例外） / NaN self-reflexive tests
          OR (fSoftLoDeg <> fSoftLoDeg) OR (fSoftHiDeg <> fSoftHiDeg)                    // 软限 NaN 判 / Soft-limit NaN tests
          OR ((fPosAct - fPosAct) <> (fPosAct - fPosAct));                                // 位置 Inf 差值自减判 / Inf test
_bCfgBad := (fSoftHiDeg <= fSoftLoDeg) OR _bNonFin;                                       // 软限几何组态闸（R151） / Soft-limit geometry gate
_bTargetBad := (fTargetDeg < (0.0 - DL_FLOAT_EPS)) OR (fTargetDeg > (DL_FULL_TURN + DL_FLOAT_EPS));   // 目标角域闸 / Target domain gate
rtExec(CLK := bExecute);                                                                  // 执行沿，每拍必调（R228A） / Execute edge
rtReset(CLK := bReset);                                                                   // 复位沿，每拍必调 / Reset edge

(* —— 段 1：单拍量预清零（锁存量不入清单，R107） —— *)
_uInfo       := 16#0000_0000;      // 信息码每拍重算 / Info recomputed every scan
bValid       := FALSE;             // 有效位每拍预清 / Valid flag preset
nErrId       := 16#0000_0000;      // 事件码缺省无事件 / Event code default none
bError       := FALSE;             // 故障标志每拍预清，故障分支同拍置位（R45 配对） / Flag preset
_bSolved     := FALSE;             // 软限求解标记预清 / Solvability marker preset

(* —— 段 2：复位沿 + 组态域闸 + 目标域闸 —— *)
IF rtReset.Q THEN                                                        // 当拍复位沿 / current-scan reset edge
    _bFault := FALSE;                                                    // 清故障锁存位（锁存量） / Clear fault latch
    _uFault := 16#0000_0000;                                             // 清故障锁存码（锁存量） / Clear latched code
    _eCause := E_DL_RspCause.eNone;                                      // 清成因（锁存量） / Clear latched cause
    IF _eState = E_DL_RspState.eFault THEN
        _eState := E_DL_RspState.eIdle;                                  // 故障相迁出唯一路径 / Sole exit from fault phase
    END_IF
END_IF
IF _bCfgBad THEN                                                         // 组态域闸 / Configuration gate
    _uFault := 16#0004_03B8;                                             // 故障级：旋转最短路径故障总码 / Fault-level: short-path fault code
    _bFault := TRUE;
    bError  := TRUE;                                                     // 故障标志同拍置位（R45 配对） / Error flag set same scan
    _eCause := E_DL_RspCause.eCfgIllegal;                                // 归因：组态非法 / Cause: illegal configuration
END_IF

(* —— 段 3：规划求解（执行沿受理；归一化走条件加减 + 迭代守卫） —— *)
IF (NOT _bFault) AND rtExec.Q THEN                                       // 执行上升沿（当拍量） / Execute rising edge
    IF _bTargetBad THEN
        _uFault := 16#0004_03B8;                                         // 故障级：目标角越域 / Fault-level: target out of domain
        _bFault := TRUE;
        bError  := TRUE;                                                 // 故障标志同拍置位（R45 配对） / Error flag set same scan
        _eCause := E_DL_RspCause.eTargetBad;                             // 归因：目标越域 / Cause: target domain
    ELSE
        _fNorm := fPosAct;                                               // 归一化起点 / Normalisation start
        _nIter := 0;                                                     // 迭代计数清零 / Clear iteration counter
        _bIterBad := FALSE;                                              // 迭代守卫标记清 / Clear guard marker
        WHILE (_fNorm >= DL_FULL_TURN) AND (_nIter < DL_ITER_MAX) DO     // 条件减（禁 MOD，R10/R48） / Conditional subtraction, no modulo
            _fNorm := _fNorm - DL_FULL_TURN;
            _nIter := _nIter + 1;                                        // 守卫计数递增 / Guard increment
        END_WHILE
        WHILE (_fNorm < 0.0) AND (_nIter < DL_ITER_MAX) DO               // 条件加（禁 MOD） / Conditional addition, no modulo
            _fNorm := _fNorm + DL_FULL_TURN;
            _nIter := _nIter + 1;
        END_WHILE
        IF _nIter >= DL_ITER_MAX THEN                                    // 超守卫：置码跳出，不死循环 / Guard tripped
            _bIterBad := TRUE;
        END_IF
        IF _bIterBad THEN
            _uFault := 16#0004_03B8;                                     // 故障级：归一化超迭代守卫 / Fault-level: iteration guard
            _bFault := TRUE;
            bError  := TRUE;
            _eCause := E_DL_RspCause.eIterGuard;                         // 归因：迭代守卫 / Cause: iteration guard
        ELSE
            _fDiff := fTargetDeg - _fNorm;                               // 最小转角候选 / Candidate shortest angle
            IF _fDiff > (DL_HALF_TURN + DL_FLOAT_EPS) THEN               // 超半圈 → 反向走短路径 / Beyond half turn, go the other way
                _fDiff := _fDiff - DL_FULL_TURN;
            ELSIF _fDiff < (0.0 - DL_HALF_TURN - DL_FLOAT_EPS) THEN      // 低于负半圈 → 正向走短路径 / Below minus half turn, go positive
                _fDiff := _fDiff + DL_FULL_TURN;
            END_IF
            IF bCwOnly AND (_fDiff < 0.0) THEN                           // 单向模式：负向改成正向等价角 / CW-only forces the positive equivalent
                _fDiff := _fDiff + DL_FULL_TURN;
            END_IF
            _fAbsCand := fPosAct + _fDiff;                               // 首选圈绝对目标位 / Preferred absolute target
            IF (_fAbsCand >= fSoftLoDeg) AND (_fAbsCand <= fSoftHiDeg) THEN
                _bSolved := TRUE;                                        // 首选圈即在软限内 / Preferred turn inside limits
            ELSE
                _fAbsCand := _fAbsCand + DL_FULL_TURN;                   // 尝试另一圈（正向一圈） / Try the next turn, positive
                IF (_fAbsCand >= fSoftLoDeg) AND (_fAbsCand <= fSoftHiDeg) THEN
                    _fDiff := _fDiff + DL_FULL_TURN;                     // 转角同步修正，保证目标位与转角自洽 / Keep angle and target consistent
                    _bSolved := TRUE;
                ELSE
                    _fAbsCand := _fAbsCand - 2.0 * DL_FULL_TURN;         // 再试另一侧（负向一圈） / Try the other turn, negative
                    IF (_fAbsCand >= fSoftLoDeg) AND (_fAbsCand <= fSoftHiDeg) THEN
                        _fDiff := _fDiff - DL_FULL_TURN;
                        _bSolved := TRUE;
                    END_IF
                END_IF
            END_IF
            IF NOT _bSolved THEN                                         // 两圈均越限：拒绝并置码 / No turn inside limits
                _uFault := 16#0004_03B8;                                 // 故障级：软限无解 / Fault-level: no solution inside limits
                _bFault := TRUE;
                bError  := TRUE;
                _eCause := E_DL_RspCause.eSoftLimit;                     // 归因：软限无解 / Cause: soft-limit no solution
            ELSE
                _fTmp := _fAbsCand;                                      // 圈号求解起点 / Turn solving start
                _nTurnCalc := 0;
                _bTurnBad := FALSE;
                WHILE (_fTmp >= DL_FULL_TURN) AND (_nTurnCalc < DL_TURN_MAX) DO
                    _fTmp := _fTmp - DL_FULL_TURN;                       // 整除点不跳圈（向量 A 已核） / Exact multiples do not skip a turn
                    _nTurnCalc := _nTurnCalc + 1;
                END_WHILE
                WHILE (_fTmp < 0.0) AND (_nTurnCalc > (0 - DL_TURN_MAX)) DO
                    _fTmp := _fTmp + DL_FULL_TURN;
                    _nTurnCalc := _nTurnCalc - 1;
                END_WHILE
                IF (_nTurnCalc >= DL_TURN_MAX) OR (_nTurnCalc <= (0 - DL_TURN_MAX)) THEN
                    _bTurnBad := TRUE;                                   // 圈号超守卫上限 / Turn guard tripped
                END_IF
                IF _bTurnBad THEN
                    _uFault := 16#0004_03B8;                             // 故障级：圈号超守卫 / Fault-level: turn guard
                    _bFault := TRUE;
                    bError  := TRUE;
                    _eCause := E_DL_RspCause.eTurnGuard;                 // 归因：圈号守卫 / Cause: turn guard
                ELSE
                    fTargetAbs := _fAbsCand;                             // 绝对目标位定稿 / Final absolute target
                    nTurnIndex := _nTurnCalc;                            // 圈号定稿 / Final turn index
                    IF _fDiff >= 0.0 THEN
                        bShortestCw := TRUE;                             // 正向（含恰好 ±180° 的正优先约定） / CW, includes the exact-half-turn convention
                    ELSE
                        bShortestCw := FALSE;                            // 反向 / CCW
                    END_IF
                    bValid := TRUE;                                      // 规划有效 / Plan valid
                    _uInfo := 16#0004_04B8;                              // 信息级：规划成功 / Info: plan succeeded
                END_IF
            END_IF
        END_IF
    END_IF
END_IF

(* —— 段 4：故障解除式（R240 全当拍量） —— *)
IF rtReset.Q AND (NOT _bCfgBad) AND (NOT _bTargetBad) AND _bSolved THEN   // 分支 1：本次复位当拍已求得软限内解 / Branch 1, solved in this very scan
    _bFault := FALSE;                                                    // 清故障锁存位（锁存量） / Clear fault latch
    _uFault := 16#0000_0000;                                             // 清故障锁存码（锁存量） / Clear latched code
    _eCause := E_DL_RspCause.eNone;                                      // 清成因（锁存量） / Clear latched cause
END_IF
IF rtReset.Q AND (NOT _bCfgBad) AND (NOT _bTargetBad)                        // 分支 2：目标角本身落在软限区间内（越限条件已解除，当拍量） / Branch 2, target angle inside limits
   AND (fTargetDeg >= fSoftLoDeg) AND (fTargetDeg <= fSoftHiDeg) THEN
    _bFault := FALSE;                                                    // 清故障锁存位（锁存量） / Clear fault latch
    _uFault := 16#0000_0000;                                             // 清故障锁存码（锁存量） / Clear latched code
    _eCause := E_DL_RspCause.eNone;                                      // 清成因（锁存量） / Clear latched cause
END_IF

(* —— 段 4A：故障锁存相位迁移闸 —— *)
IF _bFault AND (_eState <> E_DL_RspState.eFault) THEN
    _eState := E_DL_RspState.eFault;                                     // 锁存即入故障相 / Latch enters fault phase
END_IF

(* —— 段 5：相位机（ENUM 全成员显式标签 + ELSE 兜底，R128） —— *)
CASE _eState OF

E_DL_RspState.eIdle:
    IF rtExec.Q AND (NOT _bFault) THEN                                   // 出口 1：收到执行沿（结果由段 3 就地算出） / Execute edge received
        _eState := E_DL_RspState.eRun;
    ELSIF _bFault THEN                                                   // 出口 2：故障锁存 / Fault latched
        _eState := E_DL_RspState.eFault;
    END_IF

E_DL_RspState.eRun:
    IF rtReset.Q THEN                                                    // 出口 1：复位回空闲（前置消失，R98） / Reset returns idle
        _eState := E_DL_RspState.eIdle;
    ELSIF _bFault THEN                                                   // 出口 2：故障锁存 / Fault latched
        _eState := E_DL_RspState.eFault;
    END_IF

E_DL_RspState.eFault:
    ;                                                                     // 故障相：仅段 4 复位沿可迁出 / Only the reset edge leaves this phase

ELSE
    _uFault := 16#0004_03B8;                                             // 故障级：非法相位兜底（归并总码） / Illegal-phase fallback
    _bFault := TRUE;
    bError  := TRUE;
    _eCause := E_DL_RspCause.ePhaseBad;                                  // 归因：非法相位 / Cause: illegal phase
    _eState := E_DL_RspState.eFault;

END_CASE

(* —— 段 6：出口单点映射（名实同源；锁存码回放；故障相安全侧） —— *)
IF _bFault THEN
    bValid      := FALSE;                                                // 故障相规划无效 / Plan invalid in fault
    bShortestCw := FALSE;                                                // 故障相不宣称转向（保守：不给方向建议） / No direction advice in fault
    fTargetAbs  := fPosAct;                                              // 故障相目标位回落到当前位置（零位移，安全侧） / Target falls back to current position
    nTurnIndex  := 0;                                                    // 故障相圈号清零 / Turn index zeroed in fault
END_IF
IF _bFault THEN
    nErrId := _uFault;                                                   // 故障锁存码回放 / Replay latched fault code
ELSE
    nErrId := _uInfo;                                                    // 信息码 / Info code
END_IF
bError := _bFault;                                                       // 故障标志与锁存同源（名实双出口，R191） / Flag from latch
eState := _eState;                                                       // 状态出口 / State outlet
eCause := _eCause;                                                       // 成因出口 / Cause outlet

END_FUNCTION_BLOCK

(* ---- FB_DL_AxisSafetyStateMon.st ---- *)
(*
  ==================================================================
  组件名 Component  : FB_DL_AxisSafetyStateMon
  分类   Category   : DL_Motion
  复杂度 Complexity  : cx5
  版本   Version    : 1.0.0
  功能   Purpose    : 轴安全功能状态字监视。从驱动器安全状态字反馈（STO /
                      SLS / SOS 位）解码激活态，与 PLC 侧安全请求逐位比对：
                      请求-反馈不一致经消抖确认窗后锁存不一致位图并置故障
                      （仅监视不发令，无任何命令输出）；全零反馈字持续判
                      通信失效。与 AxisSs1StopSeq 执行件分工互引。
  来源   Source     : t1-6-plcopen（轴侧安全层同层扩展）
  溯源   Origin     : IEC 61131-3 标准语义的道莅防御性实现；STO / SLS / SOS
                      为 IEC 61800-5-2 公开安全功能语义，clean-room 自研实现，
                      未复制 PLCopen 或任何厂商私有库源码。
  平台   Platform   : 纯 IEC 61131-3（Standard.library: TON / R_TRIG，无私有库）
  分工声明 Split     : 与 FB_DL_AxisSs1StopSeq 分工——后者为 SS1 停车执行顺控
                      （发令侧），本件为安全功能状态字监视（收令侧仅监视，
                      零命令输出）；本件不做安全功能替代，安全回路本体仍由
                      硬件安全层承担。
  作者   Author     : 道莅代码库 · PLC 编程专家（R58）
  ------------------------------------------------------------------
  边界 Boundary     :
                      一 状态字位定义（固定掩码常量，禁变量移位 R48）：
                         位 0 = STO 激活，位 1 = SLS 激活，位 2 = SOS 激活；
                         位 3..15 保留（不参与判定，声明覆盖范围）；
                      二 不一致判据 = 请求位 XOR 反馈位逐位比对，任一位不
                         一致持续 tMismatchDebounce 后锁存位图并置故障；解除
                         路径 = bReset 上升沿（唯一路径，R188）；
                      三 通信失效判据 = 反馈字连续两拍全零且持续 tCommWatch
                         判失效（故障级独立成因，R190）；
                      四 仅监视：本件零命令输出（功能定义即不发令）；
                      五 无全局变量、无外部变量声明、无物理地址寻址。
  修订记录 Revision  :
    2026-11-21  v1.0.0  R58 首版（批 4 · 序号 13）
  ==================================================================
*)

FUNCTION_BLOCK FB_DL_AxisSafetyStateMon
VAR_INPUT
    bEnable            : BOOL := TRUE;     // 使能，失能冻结监视输出末值 [-] / enable, disabling freezes the monitor outputs
    bReset             : BOOL := FALSE;    // 复位上升沿清故障锁存 [-] / reset rising edge clears the fault latch
    bStoReq            : BOOL := FALSE;    // STO 请求（PLC 侧发出）[-] / the STO request from the PLC side
    bSlsReq            : BOOL := FALSE;    // SLS 请求 [-] / the SLS request
    bSosReq            : BOOL := FALSE;    // SOS 请求 [-] / the SOS request
    uSafFbWord         : WORD := 16#FFFF;  // 驱动器安全状态字反馈 [位图] / the drive safety status word feedback [bitmap]
    tMismatchDebounce  : TIME := T#100MS;  // 不一致消抖确认窗 [毫秒] / the mismatch debounce window [millisecond]
    tCommWatch         : TIME := T#500MS;  // 全零通信失效窗 [毫秒] / the all zero comm loss window [millisecond]
END_VAR
VAR_OUTPUT
    bStoActive : BOOL := FALSE; // STO 激活解码出口（位 0）[-] / the STO active decode outlet, bit zero
    bSlsActive : BOOL := FALSE; // SLS 激活解码出口（位 1）[-] / the SLS active decode outlet, bit one
    bSosActive : BOOL := FALSE; // SOS 激活解码出口（位 2）[-] / the SOS active decode outlet, bit two
    uMismatch  : WORD := 16#0000; // 不一致位图出口（请求 XOR 反馈，锁存回放）[位图] / the mismatch bitmap outlet, latched replay [bitmap]
    bCommBad   : BOOL := FALSE; // 通信失效指示（故障级）[-] / the comm loss indicator, fault grade
    bError     : BOOL := FALSE; // 故障锁存标志（不一致或通信失效）[-] / the fault latch flag
END_VAR
VAR
    rtReset  : R_TRIG; // 复位沿检测，段 0 无条件刷新 / the reset edge
    tonMis   : TON;    // 不一致消抖窗，段 0 无条件刷新 / the mismatch debounce window
    tonComm  : TON;    // 通信失效窗，段 0 无条件刷新 / the comm loss window
    _bStoFb  : BOOL := FALSE; // STO 反馈解码工作量（位 0）/ the STO feedback decode work bit
    _bSlsFb  : BOOL := FALSE; // SLS 反馈解码工作量（位 1）/ the SLS feedback decode work bit
    _bSosFb  : BOOL := FALSE; // SOS 反馈解码工作量（位 2）/ the SOS feedback decode work bit
    _uMisNow : WORD := 16#0000; // 当拍不一致位图工作量 [位图] / the current mismatch bitmap work value
    _bMisNow : BOOL := FALSE; // 当拍存在不一致工作量 [-] / the current mismatch work flag
    _bMisL   : BOOL := FALSE; // 不一致锁存位 [-] / the mismatch latch bit
    _uMisL   : WORD := 16#0000; // 不一致位图锁存 [位图] / the mismatch bitmap latch
    _bCommL  : BOOL := FALSE; // 通信失效锁存位 [-] / the comm loss latch bit
    _bInit   : BOOL := FALSE; // 首扫初始化完成标志（R310）/ the first scan flag
END_VAR
VAR CONSTANT
    DL_ASM_BIT_STO : WORD := 16#0001; // STO 位掩码（位 0，固定常量禁移位）/ the STO bit mask, bit zero
    DL_ASM_BIT_SLS : WORD := 16#0002; // SLS 位掩码（位 1）/ the SLS bit mask, bit one
    DL_ASM_BIT_SOS : WORD := 16#0004; // SOS 位掩码（位 2）/ the SOS bit mask, bit two
    DL_ASM_WORD_ZERO : WORD := 16#0000; // 全零字常量（通信失效判据）/ the all zero word constant
END_VAR

// 段 0｜定时器与沿检测无条件周期刷新（禁入分支，FB50-1）/ segment 0, the unconditional refresh
rtReset(CLK := bReset); // 复位沿 / the reset edge
_bStoFb := (uSafFbWord AND DL_ASM_BIT_STO) <> DL_ASM_WORD_ZERO; // 位 0 解码（固定掩码，无移位）/ the bit zero decode by a fixed mask
_bSlsFb := (uSafFbWord AND DL_ASM_BIT_SLS) <> DL_ASM_WORD_ZERO; // 位 1 解码 / the bit one decode
_bSosFb := (uSafFbWord AND DL_ASM_BIT_SOS) <> DL_ASM_WORD_ZERO; // 位 2 解码 / the bit two decode
_uMisNow := 16#0000; // 当拍位图预清零 / preset the current bitmap zero
IF bStoReq <> _bStoFb THEN // STO 请求反馈不一致 / an STO request feedback mismatch
    _uMisNow := _uMisNow OR DL_ASM_BIT_STO; // 位图记位 / mark the bitmap
END_IF
IF bSlsReq <> _bSlsFb THEN // SLS 不一致 / an SLS mismatch
    _uMisNow := _uMisNow OR DL_ASM_BIT_SLS; // 位图记位 / mark the bitmap
END_IF
IF bSosReq <> _bSosFb THEN // SOS 不一致 / an SOS mismatch
    _uMisNow := _uMisNow OR DL_ASM_BIT_SOS; // 位图记位 / mark the bitmap
END_IF
_bMisNow := _uMisNow <> DL_ASM_WORD_ZERO; // 当拍存在不一致 / a mismatch exists this scan
tonMis(IN := bEnable AND (NOT _bMisL) AND (NOT _bCommL) AND _bMisNow, PT := tMismatchDebounce); // 消抖窗，IN 串锁存反闸（防复位同拍重锁，FB50-1）/ the debounce window gated against the latches
tonComm(IN := bEnable AND (NOT _bCommL) AND (uSafFbWord = DL_ASM_WORD_ZERO), PT := tCommWatch); // 通信失效窗，IN 串全零条件 / the comm window on the all zero condition

// 段 1｜首扫初始化（R310）/ segment 1, the first scan
IF NOT _bInit THEN // 首扫一拍 / the first scan
    _bInit := TRUE; // 置首扫标志 / raise the flag
END_IF

// 段 2｜复位沿作用域：清不一致锁存与位图 / 清通信锁存 / 清出口（三项逐项声明）/ segment 2, the reset edge scope
IF rtReset.Q THEN // 复位沿 / the reset edge
    _bMisL := FALSE; // 作用域一：清不一致锁存（解除路径 = bReset 沿，R188）/ scope one, clear the mismatch latch
    _uMisL := 16#0000; // 作用域一：清位图锁存 / scope one, clear the bitmap latch
    _bCommL := FALSE; // 作用域二：清通信锁存 / scope two, clear the comm latch
    uMismatch := 16#0000; // 作用域三：清位图出口 / scope three, clear the bitmap outlet
    bCommBad := FALSE; // 作用域三：清通信出口 / scope three, clear the comm outlet
    bError := FALSE; // 作用域三：清故障出口 / scope three, clear the fault outlet
END_IF

// 段 3｜故障锁存判定（消抖确认后锁存，R190 独立成因）/ segment 3, the fault latch verdicts
IF bEnable THEN // 使能才锁存 / latch only when enabled
    IF tonMis.Q AND (NOT _bMisL) THEN // 消抖确认且未锁存 / a debounced confirmation while unlatched
        _bMisL := TRUE; // 置不一致锁存 / raise the mismatch latch
        _uMisL := _uMisNow; // 锁存首因位图（回放不重推断 R152）/ latch the first cause bitmap
    END_IF
    IF tonComm.Q AND (NOT _bCommL) THEN // 通信失效确认且未锁存 / a comm confirmation while unlatched
        _bCommL := TRUE; // 置通信锁存 / raise the comm latch
    END_IF
END_IF

// 段 4｜统一出口（边界四：仅监视，零命令输出）/ segment 4, the unified outlet
IF bEnable THEN // 使能实时刷新解码 / refresh the decode when enabled
    bStoActive := _bStoFb; // STO 出口 / the STO outlet
    bSlsActive := _bSlsFb; // SLS 出口 / the SLS outlet
    bSosActive := _bSosFb; // SOS 出口 / the SOS outlet
END_IF // 失能时解码出口冻结保持末值（R191 冻结保持声明）/ disabled freezes the decode outlets
IF _bMisL THEN // 不一致锁存回放 / the mismatch latch replay
    uMismatch := _uMisL; // 位图回放 / replay the bitmap
ELSE // 无锁存随当拍位图（信息级实时可观测）/ no latch, the live bitmap
    uMismatch := _uMisNow; // 实时位图 / the live bitmap
END_IF
bCommBad := _bCommL; // 通信出口与锁存同源 / the comm outlet shares the latch
bError := _bMisL OR _bCommL; // 故障标志聚合（R191 名实双出口）/ the flag aggregation
END_FUNCTION_BLOCK
